(* IEC 61131-3 sources: plcassist-cli/packages/volt-lsp-iec/test-corpus/pro2193/Device/Plc Logic/Application/09 Misc/Library Manager/L_TT1P_TechnologyModules (part 2) *)

(* ---- _TM_STACKERCRANEAXISCONTROLBASE.fb ---- *)
FUNCTION_BLOCK _TM_STACKERCRANEAXISCONTROLBASE EXTENDS _TM_MotionControl
VAR_OUTPUT
	PPAR : POINTER TO _scPar_TM_StackerCraneAxisControlBase;
	PSF : POINTER TO _scSF_TM_StackerCraneAxisControlBase;
	PAP : POINTER TO _scAP_TM_StackerCraneAxisControlBase;
END_VAR
VAR_IN_OUT
	AXIS : AXIS_REF;
	DATABUSIN : ITF_DataBus;
	EADDRESS : L_TT1P_StackerCraneAddress;
	LROVERRIDE : LREAL;
	XEXECUTEBRAKETEST : BOOL;
	XEXECUTEBRAKEGRINDIN : BOOL;
	XOSCCOMP : BOOL;
	LROSCCOMPPOSSCALED : LREAL;
	LROSCCOMPLOADSCALED : LREAL;
	LRACTPOS : LREAL;
	LRACTVEL : LREAL;
	XOSCCOMPACTIVE : BOOL;
	XINPOSITION : BOOL;
	XAXISREADY : BOOL;
	ECONTROLMODE : L_MC1P_ControlMode;
	XCOMMANDABORTED : BOOL;
END_VAR
VAR
	XREGULATORONINTERNAL : BOOL;
	ETMSTATE_EXITSELECTMODE : L_TT1P_States;
	XOSCCOMP_INT : BOOL;
	XOSCCOMP_OLD : BOOL;
	XEXECUTEBRAKETEST_INT : BOOL;
	XEXECUTEBRAKEGRINDIN_INT : BOOL;
	LROVERRIDE_INT : LREAL := 1;
	LRMASTERTASKCYCLETIME : LREAL;
	LRTASKCYCLETIME : LREAL;
	SCPAR_INT : _scPar_TM_StackerCraneAxisControlBase;
	EADDRESS_INT : L_TT1P_StackerCraneAddress;
	XCOMMANDABORTED_INT : BOOL;
	XDONEBRAKEGRINDIN : BOOL;
	XDONEBRAKETEST : BOOL;
	XBRAKEFUNKTIONBUSY : BOOL;
	XSTOPACTIVE_INT : BOOL;
	XJOGGINGACTIVE_INT : BOOL;
	XHOMINGACTIVE_INT : BOOL;
	XPROFILEXYBUSY_INT : BOOL;
	XPOSITIONINGBUSY_INT : BOOL;
	XPOSITIONINGDONE_INT : BOOL;
	XBRAKETESTACTIVE : BOOL;
	XBRAKEGRINDINACTIVE : BOOL;
	XOSCCOMPENABLE_INT : BOOL;
	XOSCCOMPENABLE_OLD : BOOL;
	LRTIMECOUTERCONSTANTTORQUEVALID : LREAL;
	XSTARTCONSTANTTORQUEVALID_INT : BOOL;
	LRSTARTCONSTANTTORQUE_INT : LREAL;
	LROSCCOMPPOSSCALED_INT : LREAL := 0;
	LROSCCOMPLOADSCALED_INT : LREAL := 0;
	XOSCCOMPENABLE_LOCK : BOOL;
	LROSCCOMPPOSSCALED_LOCK : LREAL;
	LROSCCOMPLOADSCALED_LOCK : LREAL;
	XUPDATEOSCCOMPPARAMETER : BOOL;
	XAMPRATIOVALID : BOOL;
	XEIGENFREQVALID : BOOL;
	WREQUESTSOSCCOMPPARMAVALID : WORD;
	WREQUESTSOSCCOMPPARMAVALID_OLD : WORD;
	XREQUESTSOSCCOMPPARMA : BOOL;
	WRTRIGOSCCOMPPARMAVALID : WORD;
	WFTRIGOSCCOMPPARMAVALID : WORD;
	XSWLIMITDISABLED : BOOL;
	XSELECTCSVACTIVE_INT : BOOL;
	XSELECTCSPACTIVE_INT : BOOL;
	XSELECTCSPBLOKEDBYOSCCOMP : BOOL;
	EAXISSTATE_OLD : L_MC1P_AXIS_STATE;
	XPOSITIONINGDONE_OLD : BOOL;
	XAXISENABLED_OLD : BOOL;
	IFOR : INT;
	XWAITNEXTCYCLEFORSETCONTROLERMODE : BOOL;
	XINPOSITIONVALID : BOOL;
	XINPOSITION_INT : BOOL;
	LRTARGETACTPOSITION : LREAL;
	LRTARGETSETPOSITION : LREAL;
	LRPOSINWINDOW : LREAL;
	LRTIMEPOSINWINDOW : LREAL := 50;
	LRACTTIMEPOSINWINDOW : LREAL;
	XHOLDPOWEROFF_INT : BOOL;
	XDISABLEAXIS_INT : BOOL;
	XDISABLEAXIS_OLD : BOOL;
	XAXISDISABLED_INT : BOOL;
	XAXISDISABLED_OLD : BOOL;
	LRTIMECOUNTER_INT : LREAL;
	WCOUNTERAXISENABLED_INT : WORD;
	WBRAKETESTMODE : WORD;
	WBRAKETESTSTEPPER : WORD;
	WBRAKEGRINDINSTEPPER : WORD;
	LRBRAKETESTCONSTANTTORQUE : LREAL;
	LRTIMECOUNTER : LREAL;
	LRTIMEBRAKERELEASE : LREAL := 0.2;
	LRTIMEIDENTTORQUE : LREAL := 0.8;
	XRESETFILTERSTANDSTILLTORQUE : BOOL;
	WBRAKEGRINDINCYCLES_INT : WORD;
	EADDRESS_LOCK : L_TT1P_StackerCraneAddress;
	XADDRESS_LOCK : BOOL;
	ECONTROLMODECAMEFROM : L_MC1P_ControlMode;
	PELEMENT : POINTER TO L_MB1P_ChannelElement;
	PRIGHT : POINTER TO L_MB1P_ChannelElement;
	PLEFT : POINTER TO L_MB1P_ChannelElement;
	PDATA : POINTER TO L_MB1P_ChannelData;
	PDATACONTROL : POINTER TO L_MB1P_ChannelData;
	PLIST : POINTER TO L_MB1P_ListControl;
	COMIN_XLOCKCOMCHANNEL : BOOL;
	COM_XENABLE : BOOL;
	COMIN_XRESETERROR_INT : BOOL;
	COMIN_XREGULATORON_INT : BOOL;
	COMIN_XSTOP_INT : BOOL;
	COMOUTTMP_WERRORID : WORD;
	COMOUTTMP_DWERRORID : DWORD;
	COMOUT_WERRORIDSTEPPER : DWORD;
	COMOUT_DWPARSTEPPER : DWORD;
	COMOUT_DWVARSTEPPER : DWORD;
	COMOUT_DWDRIVEERRORID : DWORD;
	COMOUT_XEXECUTEMOVEXY : BOOL;
	COMOUT_XEXECUTEMOVEXY_OLD : BOOL;
	WMOVEXYEXECUTESTATE : WORD;
	COMIN_XEXECUTEPROFILEXY : BOOL;
	COMIN_XMOVEXYACTIVE : BOOL;
	COMIN_XMOVEXYBUSY : BOOL;
	COMIN_XMOVEXYDONE : BOOL;
	COMIN_XMOVEXYACTIVE_OLD : BOOL;
	COMIN_XMOVEXYDONE_OLD : BOOL;
	COMIN_XMAINTENANCEMODE : BOOL;
	COMIN_XMOVEXYCOMMANDABORT : BOOL;
	COMIN_EMASTERSTATE : WORD;
	COMIN_LRSETPOSDIST : LREAL;
	COMIN_XRESETHOLDPOWEROFF : BOOL;
	FB_COMCHANNEL : L_MB1P_ComChannelSlaveState;
	XCOMMUNICATIONVALID_LOCK : BOOL;
	XERRORCOMMUNICATION : BOOL;
	XCOMMUNICATIONVALID : BOOL;
	_XCOMERRORINVALIDMASTERCONTROLMODUL : BOOL;
	_XCOMERROR : BOOL;
	_ECOMERRORID : L_IE1P_Error;
	XERROR_INVALIDSWLIMIT : BOOL;
	XERROR_INVALIDINVERTER : BOOL;
	XERROR_NOVALIDACCELERATION_MOVEABSOLUTE : BOOL;
	XERROR_INVALIDINPUT_BRAKEGRINDIN : BOOL;
	XERROR_AXISDISABLEDISREQUIRED : BOOL;
	XWARNINGCOMMUNICATION : BOOL;
	XWARNING_INVALIDINVERTER : BOOL;
	XWARNING_AXISDISABLEDISREQUIRED : BOOL;
	FB_FILTERACTSTANDSTILLTORQUE : L_USPP_PT1Filter;
	FB_FILTERACTTORQUE : L_USPP_PT1Filter;
	FB_OSCILLATIONCOMP : L_CT1P_OscillationComp;
	FB_CALCOSCILATIONCOMPPARAMETER : L_MB1P_CalcOscilationCompParameter;
	FB_SETCONTROLLERMODE : L_MC1P_SetControlMode;
	FB_BRAKETEST : L_MC1P_BrakeTest;
	FB_BRAKEGRINDIN : L_MC1P_BrakeGrindIn;
	FB_READMACHINEDATA : L_MC1P_ReadMachineData;
	FB_DISABLESWLIMIT : L_MC1P_DisableSWLimit;
	FB_WRITEBOOLPARAMETER : MC_WriteBoolParameter;
	MC_READPARAMETERPOSINWINDOW : MC_ReadParameter := STRUCT(ParameterNumber := 130);
	MC_READPARAMETERTIMEPOSINWINDOW : MC_ReadParameter := STRUCT(ParameterNumber := 131);
	FB_RESETFOLLOWINGERROR : L_MC1P_ResetFollowingError;
	MC_READPARAMETEREXTPOSITINCNTRL : MC_ReadParameter := STRUCT(ParameterNumber := 90);
	IPARFRAME : INT;
	IMAINFRAME : INT;
	IVISUTABLESETPOS : INT := 1;
END_VAR
END_FUNCTION_BLOCK

METHOD CALL_ABC
END_METHOD

METHOD CALL_ABCCTRLREQACTIVE : BOOL
END_METHOD

METHOD CALL_ABCGENERALSETTINGS
END_METHOD

METHOD CALL_ALLOCPOINTADR
END_METHOD

METHOD CALL_COMIN
END_METHOD

METHOD CALL_COMOUT
END_METHOD

METHOD CALL_CTRLREQACTIVE : BOOL
END_METHOD

METHOD CALL_ERRORHANDLER
END_METHOD

METHOD CALL_FBMETHODS
END_METHOD

METHOD CALL_FB_BRAKEGRINDIN
END_METHOD

METHOD CALL_FB_BRAKEGRINDIN_INPUT
END_METHOD

METHOD CALL_FB_BRAKETEST
END_METHOD

METHOD CALL_FB_BRAKETEST_INPUT
END_METHOD

METHOD CALL_FB_CALCOSCILATIONCOMPPARAMETER
END_METHOD

METHOD CALL_FB_CALCOSCILATIONCOMPPARAMETER_INPUT
END_METHOD

METHOD CALL_FB_COMCHANNEL
END_METHOD

METHOD CALL_FB_DISABLESWLIMIT
END_METHOD

METHOD CALL_FB_FILTERACTTORQUE
END_METHOD

METHOD CALL_FB_OSCILLATIONCOMP
END_METHOD

METHOD CALL_FB_OSCILLATIONCOMP_INPUT
END_METHOD

METHOD CALL_FB_READPARAMETERINPOSITION
END_METHOD

METHOD CALL_FB_RESETFOLLOWINGERROR
END_METHOD

METHOD CALL_FB_SETCONTROLLERMODE
END_METHOD

METHOD CALL_FB_WRITEBOOLPARAMETER
END_METHOD

METHOD CALL_INPOSITION
END_METHOD

METHOD CALL_INITDONE
END_METHOD

METHOD CALL_INITROUTINE
END_METHOD

METHOD CALL_INTERNALCTRL
END_METHOD

METHOD CALL_MOVEXYEXECUTE
END_METHOD

METHOD CALL_OUTPUT
END_METHOD

METHOD CALL_OUTPUT_SF
END_METHOD

METHOD CALL_REQUESTS_EXT
END_METHOD

METHOD CALL_RESETCOMMANDS
END_METHOD

METHOD CALL_RESETOUTPUT
END_METHOD

METHOD CALL_RESETWARNINGS
END_METHOD

METHOD CALL_STATEMACHINE
END_METHOD

METHOD CALL_STOP
END_METHOD

METHOD GET_ADDRESS : WORD
VAR_INPUT
	IELEMENTID : INT;
	EADDRESS : L_TT1P_StackerCraneAddress;
END_VAR
END_METHOD

METHOD CALL_S000_CYCLIC
END_METHOD

METHOD CALL_S002_READY
END_METHOD

METHOD CALL_S003_HOMING
END_METHOD

METHOD CALL_S010_JOGGING
END_METHOD

METHOD CALL_S014_MOVE_ABS
END_METHOD

METHOD CALL_S060_SELECTMODECSV
END_METHOD

METHOD CALL_S123_SELECTMODECSP
END_METHOD

METHOD CALL_S186_MOVE_XY
END_METHOD

METHOD CALL_S187_MAINTENANCE
END_METHOD

METHOD CALL_S188_BRAKETEST
END_METHOD

METHOD CALL_S189_BRAKEGRINDIN
END_METHOD

METHOD CALL_S996_STOP
END_METHOD

METHOD CALL_S999_ERROR
END_METHOD

METHOD CALL_T000_ALLSTATES
END_METHOD

METHOD CALL_T002_READY
END_METHOD

(* ---- _TM_STACKERCRANEHEADCONTROLBASE.fb ---- *)
FUNCTION_BLOCK _TM_STACKERCRANEHEADCONTROLBASE EXTENDS _TM_MotionControlBase
VAR_OUTPUT
	PPAR : POINTER TO _scPar_TM_StackerCraneHeadControlBase;
	PSF : POINTER TO _scSF_TM_StackerCraneHeadControlBase;
	PAP : POINTER TO _scAP_TM_StackerCraneHeadControlBase;
END_VAR
VAR_IN_OUT
	XRESETERROR : BOOL;
	XSTOPALL : BOOL;
	SCPAR : _scPar_TM_StackerCraneHeadControlBase;
	XEXECUTEPROFILEX : BOOL;
	XEXECUTEPROFILEY : BOOL;
	XMAINTENANCEMODE : BOOL;
	DATABUSOUT : ITF_DataBus;
	XAXESREADY : BOOL;
	XAXESENABLED : BOOL;
	SCSIGNALFLOW : _scSF_TM_StackerCraneHeadControlBase;
	XAXESHOMED : BOOL;
	XPROFILEXDONE : BOOL;
	XPROFILEYDONE : BOOL;
	XPROFILEXBUSY : BOOL;
	XPROFILEYBUSY : BOOL;
	XERROR : BOOL;
	XWARNING : BOOL;
	EERRORID : L_IE1P_Error;
	ASCERRORINFO : ARRAY [1..6] OF L_TT1P_scErrorInfo;
END_VAR
VAR
	AXDONENEXTCYCLE_INT : ARRAY [1..2] OF BOOL;
	ADWREQUESTSINFOCOMIN : ARRAY [1..2] OF DWORD;
	ADWREQUESTSINFOCOMIN_OLD : ARRAY [1..2] OF DWORD;
	ADWFTRIGCOMIN : ARRAY [1..2] OF DWORD;
	ADWRTRIGCOMIN : ARRAY [1..2] OF DWORD;
	LRMASTERTASKCYCLETIME : LREAL;
	LRTASKCYCLETIME : LREAL;
	SCPAR_INT : _scPar_TM_StackerCraneHeadControlBase;
	XEXECUTEPROFILEX_INT : BOOL;
	XEXECUTEPROFILEY_INT : BOOL;
	XSTOPALL_INT : BOOL;
	XMAINTENANCEMODE_INT : BOOL;
	AXPOSITIONINGDONE_INT : ARRAY [1..2] OF BOOL;
	XPOSITIONINGDONE_INT : BOOL;
	XPOSITIONINGBUSY_INT : BOOL;
	IWAITTASKCYCLESFROSTATUSFORMCOM_INT : LREAL := 100;
	AICOUNTTASKCYCLES_INT : ARRAY [1..c_iNumOfAxisModule] OF INT;
	XXYCONTROLLERWAITSTARTX_INT : BOOL;
	XXYCONTROLLERWAITSTARTY_INT : BOOL;
	XCOMMUNICATIONVALID : BOOL;
	XLOCKCOMCHANNEL : BOOL;
	IFOR : INT;
	IDX1 : INT;
	WTEMP : WORD;
	DWTEMP : DWORD;
	DWTEMP1 : DWORD;
	DWSTATUSWORDTEMP : DWORD;
	COMIN_AXISIDX : INT;
	XWAITSTARTX_OLD : BOOL;
	XWAITSTARTY_OLD : BOOL;
	XPROFILEEXECUTE1X_OLD : BOOL;
	XPROFILEEXECUTE1Y_OLD : BOOL;
	XPROFILEEXECUTE2X_OLD : BOOL;
	XPROFILEEXECUTE2Y_OLD : BOOL;
	PLIST : POINTER TO L_MB1P_ListControl;
	PELEMENT : POINTER TO L_MB1P_ChannelElement;
	PDATA : POINTER TO L_MB1P_ChannelData;
	PDATA_AXISX : POINTER TO L_MB1P_ChannelData;
	PDATA_AXISY : POINTER TO L_MB1P_ChannelData;
	PRIGHT : POINTER TO L_MB1P_ChannelElement;
	PLEFT : POINTER TO L_MB1P_ChannelElement;
	COM_XENABLE : BOOL;
	COMIN_INUMOFAXES : INT;
	COMIN_XLOCKCOMCHANNEL : BOOL;
	COMIN_XXAXISCONTROLAVAILABLE : BOOL;
	COMIN_XYAXISCONTROLAVAILABLE : BOOL;
	COMIN_XAPAXISCONTROLAVAILABLE : BOOL;
	COMIN_XSLAVEXAXISCONTROLAVAILABLE : BOOL;
	COMIN_XSLAVEYAXISCONTROLAVAILABLE : BOOL;
	COMIN_XPOINTERTOXAXISVALID : BOOL;
	COMIN_AWPARVALIDMASK : ARRAY [1..6] OF WORD;
	COMIN_AXAXISVALID : ARRAY [1..c_iNumOfAxisModule] OF BOOL;
	COMIN_XAXESENABLED : BOOL;
	COMIN_XAXESREADY : BOOL;
	COMIN_XAXESHOMED : BOOL;
	COMIN_XSTOP : BOOL;
	COMIN_AXAXISREADY : ARRAY [1..c_iNumOfAxisModule] OF BOOL;
	COMIN_AXAXISENABLED : ARRAY [1..c_iNumOfAxisModule] OF BOOL;
	COMIN_AXHOMINGBUSY : ARRAY [1..c_iNumOfAxisModule] OF BOOL;
	COMIN_AXISHOMED : ARRAY [1..c_iNumOfAxisModule] OF BOOL;
	COMIN_AXSTOPACTIVE : ARRAY [1..c_iNumOfAxisModule] OF BOOL;
	COMIN_AXERROR : ARRAY [1..c_iNumOfAxisModule] OF BOOL;
	COMIN_AXWARNING : ARRAY [1..c_iNumOfAxisModule] OF BOOL;
	COMIN_AXABCCTRLREQACTIVE : ARRAY [1..c_iNumOfAxisModule] OF BOOL;
	COMIN_AXINPOSITION : ARRAY [1..c_iNumOfAxisModule] OF BOOL;
	COMIN_AETMSTATE : ARRAY [1..c_iNumOfAxisModule] OF WORD;
	COMIN_EERRORID : WORD;
	COMIN_AEERRORID : ARRAY [1..c_iNumOfAxisModule] OF WORD;
	COMIN_ASCERRORINFO : ARRAY [1..c_iNumOfAxisModule] OF L_TT1P_scErrorInfo;
	COMIN_AXXYPROFILEBUSY : ARRAY [1..c_iNumOfAxisModule] OF BOOL;
	COMIN_AXPOSITIONINGBUSY : ARRAY [1..c_iNumOfAxisModule] OF BOOL;
	COMIN_AXPOSITIONINGDONE : ARRAY [1..c_iNumOfAxisModule] OF BOOL;
	COMIN_ASCMINLIMITS : ARRAY [1..c_iNumOfAxisModule] OF L_TT1P_XYLimits;
	COMIN_ALRBUFFERPOSITIONNEG : ARRAY [1..c_iNumOfAxisModule] OF LREAL;
	COMIN_ALRBUFFERPOSITIONPOS : ARRAY [1..c_iNumOfAxisModule] OF LREAL;
	COMIN_ALRBUFFERVELNEG : ARRAY [1..c_iNumOfAxisModule] OF LREAL;
	COMIN_ALRBUFFERVELPOS : ARRAY [1..c_iNumOfAxisModule] OF LREAL;
	COMIN_AXBUFFERRANGE : ARRAY [1..c_iNumOfAxisModule] OF BOOL;
	COMIN_AXEXECUTEMOVEXY : ARRAY [1..c_iNumOfAxisModule] OF BOOL;
	COMIN_AXEXECUTEMOVEXY_OLD : ARRAY [1..c_iNumOfAxisModule] OF BOOL;
	COMIN_AXHOLDPOWEROFF : ARRAY [1..c_iNumOfAxisModule] OF BOOL;
	COMIN_AXPAXISVALID : ARRAY [1..c_iNumOfAxisModule] OF BOOL;
	COMIN_APAXIS : ARRAY [1..c_iNumOfAxisModule] OF POINTER TO AXIS_REF;
	COMOUT_AXRESETHOLDPOWEROFF : ARRAY [1..c_iNumOfAxisModule] OF BOOL;
	COMIN_AXOSCACTIVE : ARRAY [1..c_iNumOfAxisModule] OF BOOL;
	COMIN_AXBRAKETESTBUSY : ARRAY [1..c_iNumOfAxisModule] OF BOOL;
	COMIN_AXBRAKETESTDONE : ARRAY [1..c_iNumOfAxisModule] OF BOOL;
	COMIN_AXBRAKEGRINDINBUSY : ARRAY [1..c_iNumOfAxisModule] OF BOOL;
	COMIN_AXBRAKEGRINDINDONE : ARRAY [1..c_iNumOfAxisModule] OF BOOL;
	COMOUT_XEXECUTEPROFILEX_INT : BOOL;
	COMOUT_XEXECUTEPROFILEY_INT : BOOL;
	FB_COMCHANNEL : L_MB1P_ComChannelState;
	COMIN_XERROR_NOSTACKERCRANEAXIS : BOOL;
	XCOMMUNICATIONVALID_LOCK : BOOL;
	XERRORCOMMUNICATION : BOOL;
	_XCOMERRORINVALIDMASTERCONTROLMODUL : BOOL;
	_XCOMERROR : BOOL;
	_ECOMERRORID : L_IE1P_Error;
	XERRORDUPLICATEDADDRESS : BOOL;
	XWARNINGCOMMUNICATION : BOOL;
	XWARNING_EXECUTEXNOTPOSSIBLE : BOOL;
	XWARNING_EXECUTEYNOTPOSSIBLE : BOOL;
	XWARNING_XAXISINSERVICE : BOOL;
	XWARNING_YAXISINSERVICE : BOOL;
	XWARNING_XAXISENABLEDREQUIRED : BOOL;
	XWARNING_YAXISENABLEDREQUIRED : BOOL;
	PXAXIS : POINTER TO AXIS_REF;
	PYAXIS : POINTER TO AXIS_REF;
	XEXECUTEX_INT : BOOL;
	XEXECUTEY_INT : BOOL;
	XXYCONTROLLER_REEXECUTEX : BOOL;
	XXYCONTROLLER_REEXECUTEY : BOOL;
	EPROFILEMODEX_INT : L_TT1P_XYProfileMode;
	EPROFILEMODEY_INT : L_TT1P_XYProfileMode;
	FB_XYCONTROLLER : L_TF1P_XYController;
	IPARFRAME : INT;
	IMAINFRAME : INT;
	IVISUSELECTAXIS : INT := 1;
	ASTVISUSELECTAXIS : ARRAY [0..6] OF STRING := ['no axis selected', 'AxisX', 'AxisY', 'SlaveAxisX', 'SlaveAxisY', 'AntiPendlum', 'free axis'];
	C_INUMOFAXISMODULE : INT := 6;
END_VAR
END_FUNCTION_BLOCK

METHOD CALL_ABCCTRLREQACTIVE : BOOL
END_METHOD

METHOD CALL_ALLOCPOINTADR
END_METHOD

METHOD CALL_CHECKREQUESTS
END_METHOD

METHOD CALL_COMCHANNEL_MOVEXY
END_METHOD

METHOD CALL_COMIN
END_METHOD

METHOD CALL_COMOUT
END_METHOD

METHOD CALL_COMOUT_XYCONTROLLER_EXECUTE
END_METHOD

METHOD CALL_ERRORHANDLER
END_METHOD

METHOD CALL_ERRORHANDLER_SCERRORINFO
END_METHOD

METHOD CALL_FBMETHODS
END_METHOD

METHOD CALL_FB_COMCHANNEL
END_METHOD

METHOD CALL_FB_XYCONTROLLER
END_METHOD

METHOD CALL_FB_XYCONTROLLER_INPUT
END_METHOD

METHOD CALL_INITDONE
END_METHOD

METHOD CALL_INITROUTINE
END_METHOD

METHOD CALL_INTERNALCTRL
END_METHOD

METHOD CALL_OUTPUT
END_METHOD

METHOD CALL_OUTPUT_SF
END_METHOD

METHOD CALL_REQUESTS_COMIN
END_METHOD

METHOD CALL_REQUESTS_EXT
END_METHOD

METHOD CALL_RESETCOMMANDS
END_METHOD

METHOD CALL_RESETCOUNTER
END_METHOD

METHOD CALL_RESETOUTPUT
END_METHOD

METHOD CALL_RESETWARNINGS
END_METHOD

METHOD CALL_STATEMACHINE
END_METHOD

METHOD CALL_TMFUNCTIONALITY
END_METHOD

METHOD CALL_S000_CYCLIC
END_METHOD

METHOD CALL_S002_READY
END_METHOD

METHOD CALL_S186_MOVE_XY
END_METHOD

METHOD CALL_S187_MAINTENANCE
END_METHOD

METHOD CALL_S996_STOP
END_METHOD

METHOD CALL_S998_SERVICE
END_METHOD

METHOD CALL_S999_ERROR
END_METHOD

METHOD CALL_T000_ALLSTATES
END_METHOD

METHOD CALL_T002_READY
END_METHOD

(* ---- _TM_TABLEPOSITIONINGBASE.fb ---- *)
FUNCTION_BLOCK _TM_TABLEPOSITIONINGBASE EXTENDS _TM_MotionControl
VAR_OUTPUT
	PPAR : POINTER TO _scPar_TM_TablePositioningHigh;
	PSF : POINTER TO _scSF_TM_TablePositioningHigh;
	PAP : POINTER TO _scSF_TM_TablePositioningHigh;
END_VAR
VAR_IN_OUT
	AXIS : AXIS_REF;
	XRESETHOMEPOSITION : BOOL;
	XHWLIMITPOS : BOOL;
	XHWLIMITNEG : BOOL;
	XEXECUTEPOSITIONING : BOOL;
	XABORTPOSITIONING : BOOL;
	XFINISHPOSITIONING : BOOL;
	EPROFILENUMBER : L_TT1P_ProfileNumber;
	XTPRECEIVE : BOOL;
	LRACTTPPOSITION : LREAL;
	LRCYCPOSEXTENCODER : LREAL;
	LRSETTORQUELIMITPOS : LREAL;
	LRSETTORQUELIMITNEG : LREAL;
	LRSETOVERRIDEVELOCITY : LREAL;
	LRSETOVERRIDEACCDEC : LREAL;
	LRSETOVERRIDEJERK : LREAL;
	XPOSITIONINGACTIVE : BOOL;
	XPOSITIONINGDONE : BOOL;
	XDRIVEINTARGET : BOOL;
	LRACTPOS : LREAL;
	LRACTVEL : LREAL;
	LRACTFOLLOWINGERROR : LREAL;
	XTPRECEIVED : BOOL;
	XTPMISSED : BOOL;
	XTPOUTOFWINDOW : BOOL;
	EACTIVEPROFILE : L_TT1P_ProfileNumber;
END_VAR
VAR
	SCPAR_INT : _scPar_TM_TablePositioningHigh;
	XEXECUTEPOSITIONING_INT : BOOL;
	XABORTPOSITIONING_INT : BOOL;
	XFINISHPOSITIONING_INT : BOOL;
	XAUTOMATICUPDATE_INT : BOOL;
	LRACTTPPOSITION_INT : LREAL;
	EPROFILENUMBER_INT : L_TT1P_ProfileNumber;
	LRSETTORQUELIMITPOS_INT : LREAL;
	LRSETTORQUELIMITNEG_INT : LREAL;
	LRSETOVERRIDEVELOCITY_INT : LREAL;
	LRSETOVERRIDEACCDEC_INT : LREAL;
	LRSETOVERRIDEJERK_INT : LREAL;
	XRESETHOMEPOSITION_INT : BOOL;
	XHWLIMITPOS_INT : BOOL;
	XHWLIMITNEG_INT : BOOL;
	XTPRECEIVED_INT : BOOL;
	XTPMISSED_INT : BOOL;
	XTPOUTOFWINDOW_INT : BOOL := FALSE;
	XPOSITIONINGACTIVE_INT : BOOL;
	XPOSITIONINGDONE_INT : BOOL;
	XTPRECEIVE_INT : BOOL := FALSE;
	BYSTEPPER : BYTE;
	WSEQUENCEPROFILE : WORD := 0;
	XSEQUENCEPROFILEACTIVE : BOOL;
	XPOSDISABLEFOLLOWPROFILE : BOOL;
	LRSETPOSSEQUENCEPROFILE : LREAL;
	LRSETPOSFINISHTARGET : LREAL;
	LRFINALPOSITION : LREAL;
	XINTARGET : BOOL;
	XHOMINGEXECUTEOLD_INT : BOOL;
	HWLIMITSWITCHINTERFACE : L_MC1P_HWLimitSwitchInterface;
	RESETHOMEPOSITION : L_MC1P_ResetHomePosition;
	SMC_MOVECONTINUOUSABSOLUTE : MC_MoveContinuousAbsolute;
	SMC_MOVECONTINUOUSRELATIVE : MC_MoveContinuousRelative;
	TORQUELIMITS : L_MC1P_SetTorqueLimit;
	MC_HALT : MC_Halt;
	CONVERTTP : L_MB1P_TpConvertTp;
	READWINDOWPARAMETER : MC_ReadParameter;
	LRTARGETDISTANCE_INT : LREAL := 0;
	XPOSITIONINGABORTED_INT : BOOL := FALSE;
	XTPINSIDEWINDOW : BOOL := FALSE;
	LRTPPOSITIONINGTARGET : LREAL;
	LRACTUALPROFILEDISTANCE : LREAL;
	LRPOSITIONOLD : LREAL;
	XRESTARTPROFILE : BOOL;
	WCOUNTER : WORD;
	XEXECUTEOLD : BOOL;
	LRVELOCITYOLD : LREAL;
	XSTARTPROFILEOLD : BOOL;
	XRESTARTVELPROFILE : BOOL;
	XERRORTRAVERSIONRANGE : BOOL := FALSE;
	XNOPROFILESELECTED : BOOL := FALSE;
	XPOSITIONINGMODEINVALID : BOOL := FALSE;
	XAXISNOTHOMED : BOOL := FALSE;
	XTPRECEIVEOLD : BOOL := FALSE;
	EABORTEDPROFILE : L_TT1P_ProfileNumber;
	XTPWINDOWOPEN : BOOL;
	LRFINALPOSITIONMODULO : LREAL;
	XVISPOINTMIN : BOOL;
	XVISPOINTMAX : BOOL;
	XVISUSETPOSUP : BOOL;
	XVISUSETPOSDOWN : BOOL;
	RTRIGUP : R_TRIG;
	RTRIGDOWN : R_TRIG;
	IMAXPOINTS : INT := 13;
	IPOINT : INT := 1;
	LRTARGETWINDOW : LREAL;
	XINSIDEWINDOWFLAG : BOOL;
	XTPOUTSIDEWINDOW_TPMETHOD : BOOL;
	XTPINSIDEWINDOW_TPMETHOD : BOOL;
	LRACTUALSEQUENCESTARTPOSITION : LREAL;
	XPROFILECHAININGWITHVELOCITY : BOOL;
	XTPOUTSIDEOFWINDOW : BOOL := FALSE;
	PXMOVEFUNBUSY : POINTER TO BOOL;
	ISTATESTEPPER : INT := 0;
	XFIRSTPOSITIONINGCYCLE : BOOL := TRUE;
	XAXISVIRTUAL : BOOL := FALSE;
	XINENDVELOCITY : BOOL := FALSE;
	XTPPROFILEACTIVE : BOOL;
	XTPDURINGPOSITIONING : BOOL := FALSE;
	XPOSITIVEPROFILEVELOCITY : BOOL;
	XABORTACTIVE_INT : BOOL;
	XFINISHINGPOSITIONING_INT : BOOL;
	XEXECUTEPOSITIONINGFLAG : BOOL;
	XFINISHPOSITIONINGFLAG : BOOL;
	XABSOLUTEINENDVELOCITYOLD : BOOL;
	XRELATIVEINENDVELOCITYOLD : BOOL;
	XFUNDONEOLD : BOOL;
	XINPOSITIONOLD : BOOL;
	XFUNBUSYOLD : BOOL := FALSE;
	XPOSITIONINGDONEACTIVE : BOOL := FALSE;
	XABORTBUSYOLD : BOOL := FALSE;
	LRSETPOSITIONOLD : LREAL;
	XLASTPROFILE : BOOL;
	XCINHNOERROR : BOOL := FALSE;
	LRMODULOTARGETPOS : LREAL := 0;
	LRDIFFINSIDECYCLE : LREAL := 0;
	LRINTEGRATOR : LREAL;
	XINTEGRATORACTIVE : BOOL;
	XMOVERELEXECUTEOLD : BOOL;
	XEXECUTEMOVECONTINUOUSOLD : BOOL;
	XFIRSTSTARTRELATIVEPROFILE : BOOL;
END_VAR
END_FUNCTION_BLOCK

METHOD CALL_MC_SETTORQUE_INPUT
END_METHOD

METHOD CALL_ALLOCPOINTADR
END_METHOD

METHOD CALL_ERRORHANDLER
END_METHOD

METHOD CALL_FBMETHODS
END_METHOD

METHOD CALL_FBS
END_METHOD

METHOD CALL_FIRSTCYCLE
END_METHOD

METHOD CALL_INITDONE
END_METHOD

METHOD CALL_INITROUTINE
END_METHOD

METHOD CALL_INTERNALCTRL
END_METHOD

METHOD CALL_MC1P_HWLIMITSWITCH
END_METHOD

METHOD CALL_MC1P_RESETHOMEPOSITION
END_METHOD

METHOD CALL_OUTPUT
END_METHOD

METHOD CALL_READPOSITIONINGWINDOW
END_METHOD

METHOD CALL_REQUESTS_EXT
END_METHOD

METHOD CALL_RESETCOMMANDS
END_METHOD

METHOD CALL_RESETOUTPUTS
END_METHOD

METHOD CALL_STATEMACHINE
END_METHOD

METHOD CALL_TOUCHPROBESOURCE
END_METHOD

METHOD CALL_TPWINDOWSTATUS
END_METHOD

METHOD CALL_VISUPROFILES
END_METHOD

METHOD CALL_ABC
END_METHOD

METHOD CALL_020_RELATIVEENTRY
END_METHOD

METHOD CALL_022_RELATIVEFINALVELOCITY
END_METHOD

METHOD CALL_024_RELATIVE
END_METHOD

METHOD CALL_02_STARTSEQUENCEPROFILES
END_METHOD

METHOD CALL_110_ABORTPOSITIONING
END_METHOD

METHOD CALL_200_ERROR
END_METHOD

METHOD CALL_90_SEQUENCEPROFILE
END_METHOD

METHOD CALL_S000_CYCLIC
END_METHOD

METHOD CALL_S080_POSITIONING
END_METHOD

METHOD CALL_S081_POSITIONING_EXIT
END_METHOD

METHOD CALL_S996_STOP
END_METHOD

METHOD CALL_S999_ERROR
END_METHOD

METHOD CALL_T002_READY
END_METHOD

(* ---- _TM_VIRTUALMASTERBASE.fb ---- *)
FUNCTION_BLOCK _TM_VIRTUALMASTERBASE EXTENDS _TM_MotionControl
VAR_OUTPUT
	PPAR : POINTER TO _scPar_TM_VirtualMasterHigh;
END_VAR
VAR_IN_OUT
	VIRTUALAXIS : AXIS_REF;
	XCONTINUOUS : BOOL;
	XCYCLE : BOOL;
	XLOADSTARTPOS : BOOL;
	LRSETVEL : LREAL;
	LRSTARTPOS : LREAL;
	LRTARGETPOS : LREAL;
	XINTARGET : BOOL;
	LRACTPOS : LREAL;
	LRACTVEL : LREAL;
	LRSETPOSOUT : LREAL;
	LRSETVELOUT : LREAL;
END_VAR
VAR
	SCPAR_INT : _scPar_TM_VirtualMasterHigh;
	XCONTINUOUS_INT : BOOL;
	XCYCLE_INT : BOOL;
	XLOADSTARTPOS_INT : BOOL;
	LRSTARTPOS_INT : LREAL;
	LRTARGETPOS_INT : LREAL;
	LRSETVEL_INT : LREAL;
	LRSETVEL_LOCK : LREAL;
	EDIRECTION_LOCK : MC_DIRECTION;
	XSYNCMASTERAXIS_INT : BOOL;
	LRMASTERSTARTDISTANCE_INT : LREAL;
	LRMASTERSYNCPOSITION_INT : LREAL;
	LRSLAVESYNCPOSITION_INT : LREAL;
	WOLDSTATE : WORD;
	XSYNCMASTERAXIS_OLD : BOOL;
	XCONTINUOUS_OLD : BOOL;
	XCYCLE_OLD : BOOL;
	XSTOP_OLD : BOOL;
	XLOADSTARTPOS_OLD : BOOL;
	XOLDENABLE : BOOL;
	XSTARTPOSOUTRANGE : BOOL;
	LRTARGETPOS_SAVE : LREAL;
	XSP_EXECUTE : BOOL;
	XSP_STARTED : BOOL;
	XMOVETOTARGETPOSACTIVE : BOOL;
	BYSTEPPERMOVETOTARGETPOS : BYTE;
	LRCYCLELENGTH : LREAL;
	XMASTERITFVALID : BOOL;
	BYMASTERID : POINTER TO BYTE;
	XMASTERITFVALID_LOCK : BOOL;
	BYMASTERID_LOCK : POINTER TO BYTE;
	EMASTERTRAVERSINGRANGE : L_MC1P_TraversingRange;
	LRMASTERCYCLELENGTH : LREAL;
	LRMASTERSETPOSITIONFORSYNC : LREAL;
	LRMASTERSETVELOCITYFORSYNC : LREAL;
	LRMASTERSETACCELERATIONFORSYNC : LREAL;
	XSYNCOUTATTARGETPOS : BOOL;
	XSYNCOUTATTARGETPOSACTIVE : BOOL;
	XINTERNALCONTR_R_EDGE : R_TRIG;
	FB_SETPOSITION : MC_SetPosition;
END_VAR
END_FUNCTION_BLOCK

METHOD CALL_ABC
END_METHOD

METHOD CALL_ALLOCPOINTADR
END_METHOD

METHOD CALL_ERRORHANDLER
END_METHOD

METHOD CALL_FBMETHODS
END_METHOD

METHOD CALL_INITROUTINE
END_METHOD

METHOD CALL_INTERNALCTRL
END_METHOD

METHOD CALL_MC_SETPOSITION
END_METHOD

METHOD CALL_MASTERAXISREF
VAR_INPUT
	MASTERAXIS : L_MC1P_IAXIS_REF_MASTERVALUES;
END_VAR
END_METHOD

METHOD CALL_OUTPUT
END_METHOD

METHOD CALL_REQUESTS_EXT
END_METHOD

METHOD CALL_RESETABCMOVEEXECUTE
END_METHOD

METHOD CALL_RESETCOMMANDS
END_METHOD

METHOD CALL_RESETOUTPUT
END_METHOD

METHOD CALL_SETABCMOVEPAR
END_METHOD

METHOD CALL_SETABCMOVESETVEL
END_METHOD

METHOD CALL_STATEMACHINE
END_METHOD

METHOD CALL_S000_CYCLIC
END_METHOD

METHOD CALL_S002_READY
END_METHOD

METHOD CALL_S035_MOVE_TO_TARGET_POS
END_METHOD

METHOD CALL_S060_CONTMOTION
END_METHOD

METHOD CALL_S130_CYCLICMOTION
END_METHOD

METHOD CALL_S999_ERROR
END_METHOD

METHOD CALL_T002_READY
END_METHOD

METHOD CALL_T035_MOVE_TO_TARGET_POS
END_METHOD

METHOD CALL_T060_CONTMOTION
END_METHOD

(* ---- _TM_VIRTUALMASTERHIGH.fb ---- *)
FUNCTION_BLOCK _TM_VIRTUALMASTERHIGH EXTENDS _TM_VirtualMasterBase
VAR_INPUT
	MASTERAXIS : L_MC1P_IAXIS_REF_MASTERVALUES;
END_VAR
VAR_IN_OUT
	XSYNCMASTERAXIS : BOOL;
	XACCDECSYNC : BOOL;
	XSYNCHRONISED : BOOL;
END_VAR
VAR
	XWARNING_SYNCMODEVELACCREQUIRED : BOOL;
	XWARNING_INVALIDSYNCSLAVEDIRECTION : BOOL;
	XERROR_INVALIDSYNCSLAVEDIRECTION : BOOL;
	BYSTEPPESYNCOUTATTARGETPOS : BYTE;
	XCONTMOTION2SYNC : BOOL;
	XMOVETARGET2CONTMOTION : BOOL;
	FB_CLUTCHEXTENDEDBASE : L_MB1P_ClutchExtendedBase;
	FB_AXISCONTROLBYPOS : L_MC1P_ControlSetValues;
END_VAR
END_FUNCTION_BLOCK

METHOD CALL_ERRORHANDLER
END_METHOD

METHOD CALL_FBMETHODS
END_METHOD

METHOD CALL_FB_AXISCONTROLBYPOS
END_METHOD

METHOD CALL_FB_CLUTCHEXTENDEDBASE
END_METHOD

METHOD CALL_INITROUTINE
END_METHOD

METHOD CALL_INTERNALCTRL
END_METHOD

METHOD CALL_INTERNALCTRLSTATE
END_METHOD

METHOD CALL_OUTPUT
END_METHOD

METHOD CALL_REQUESTS_EXT
END_METHOD

METHOD CALL_RESETCOMMANDS
END_METHOD

METHOD CALL_SETCLUTCHPOSPAR
END_METHOD

METHOD CALL_STATEMACHINE
END_METHOD

METHOD CALL_SYNCDRIVE
END_METHOD

METHOD SWITCHTOEXTMASTER
END_METHOD

METHOD CALL_S030_SYNCHRONISING_POS
END_METHOD

METHOD CALL_S031_POS_IS_SYNCHRONISED
END_METHOD

METHOD CALL_S035_MOVE_TO_TARGET_POS
END_METHOD

METHOD CALL_S060_CONTMOTION
END_METHOD

METHOD CALL_S999_ERROR
END_METHOD

METHOD CALL_T002_READY
END_METHOD

METHOD CALL_T035_MOVE_TO_TARGET_POS
END_METHOD

METHOD CALL_T060_CONTMOTION
END_METHOD

(* ---- _TM_VIRTUALMASTERSTATE.fb ---- *)
FUNCTION_BLOCK _TM_VIRTUALMASTERSTATE EXTENDS _TM_VirtualMasterBase
VAR_INPUT
	MASTERAXIS : L_MC1P_IAXIS_REF_MASTERVALUES;
END_VAR
VAR_OUTPUT
	PPARSTATE : POINTER TO _scPar_TM_VirtualMasterStateExtension;
END_VAR
VAR_IN_OUT
	XSYNCMASTERAXIS : BOOL;
	XACCDECSYNC : BOOL;
	XSYNCHRONISED : BOOL;
END_VAR
VAR
	SCPARSTATE_INT : _scPar_TM_VirtualMasterStateExtension;
	GEARIN : MC_GearIn;
END_VAR
END_FUNCTION_BLOCK

METHOD CALL_ALLOCPOINTADR
END_METHOD

METHOD CALL_ALLOCPOINTADRSTATE
END_METHOD

METHOD CALL_ERRORHANDLER
END_METHOD

METHOD CALL_FBMETHODS
END_METHOD

METHOD CALL_GEARIN
END_METHOD

METHOD CALL_INITROUTINE
END_METHOD

METHOD CALL_INTERNALCTRL
END_METHOD

METHOD CALL_INTERNALCTRLSTATE
END_METHOD

METHOD CALL_OUTPUT
END_METHOD

METHOD CALL_RESETCOMMANDS
END_METHOD

METHOD CALL_RESETOUTPUT
END_METHOD

METHOD CALL_STATEMACHINE
END_METHOD

METHOD SWITCHTOEXTMASTER
END_METHOD

METHOD CALL_S000_CYCLIC
END_METHOD

METHOD CALL_S040_SYNCHRONISING_VEL
END_METHOD

METHOD CALL_S041_VELSYNCHRONISED
END_METHOD

METHOD CALL_S999_ERROR
END_METHOD

(* ---- _TM_WINDER.fb ---- *)
FUNCTION_BLOCK _TM_WINDER EXTENDS _TM_MotionControl
VAR_IN_OUT
	AXIS : AXIS_REF;
	MATERIALCOUNTERAXIS : L_MC1P_IAXIS_REF_POOL;
	PERSISTENTVAR : L_TT1P_PersistentVarWinder;
	XMATERIALFEEDING : BOOL;
	XWINDINGDIRECTION : BOOL;
	XLOADDIAM : BOOL;
	LRSETDIAM : LREAL;
	XHOLDDIAM : BOOL;
	XDIAMCALCREDUCED : BOOL;
	XWEBBREAKMONIT : BOOL;
	XJOGLINEPOS : BOOL;
	XJOGLINENEG : BOOL;
	XTRIMLINEPOS : BOOL;
	XTRIMLINENEG : BOOL;
	XSYNCLINEVEL : BOOL;
	XTENSCURVE : BOOL;
	LRSETTENS : LREAL;
	LRSETLINEVEL : LREAL;
	XSETMATERIALCOUNTER : BOOL;
	XSYNCHRONISED : BOOL;
	XACCDECSYNC : BOOL;
	XUNWIND : BOOL;
	XWEBBREAK : BOOL;
	XHOLDDIAMACTIVE : BOOL;
	XDIAMMAX : BOOL;
	XDIAMMIN : BOOL;
	LRSETDIAMOUT : LREAL;
	LRSETDIAMSCALEDOUT : LREAL;
	LRSETLINEVELSCALEDOUT : LREAL;
	LRACTTOTALTRQSCALED : LREAL;
	LRWNDSPDREF : LREAL;
	LRMATERIALCOUNTER : LREAL;
	LRLIMITLINEVEL : LREAL;
END_VAR
VAR
	XWINDINGDIRECTION_INT : BOOL := FALSE;
	XWINDINGDIRECTIONSTANDSTILL_INT : BOOL := FALSE;
	XMATERIALFEEDING_INT : BOOL := FALSE;
	XLOADDIAM_INT : BOOL;
	LRSETDIAM_INT : LREAL;
	XHOLDDIAM_INT : BOOL;
	XDIAMCALCREDUCED_INT : BOOL;
	XWEBBREAKMONIT_INT : BOOL;
	XJOGLINEPOS_INT : BOOL;
	XJOGLINENEG_INT : BOOL;
	XTRIMLINEPOS_INT : BOOL;
	XTRIMLINENEG_INT : BOOL;
	XSYNCLINEVEL_INT : BOOL;
	LRSETTENS_INT : LREAL;
	XTENSCURVE_INT : BOOL;
	XSYNCHRONISED_INT : BOOL;
	XACCDECSYNC_INT : BOOL;
	XSETMATERIALCOUNTER_INT : BOOL;
	AP10_XSETTRQOFFSET_INT : BOOL;
	AP10_LRSETTRQOFFSET_INT : LREAL;
	AP09_XSETVELOFFSET_INT : BOOL;
	AP09_LRSETVELOFFSET_INT : LREAL;
	XLINEVELDIAMCALC_INT : BOOL;
	LRSETLINEVELDIAMCALC_INT : LREAL;
	XSYNCLINEVEL_INT_OLD : BOOL;
	XUNWIND_OLD : BOOL;
	LRSETDIAMOUT_OLD : LREAL;
	XLOADDIAM_INT_OLD : BOOL;
	XERRORINVALIDINVERTER : BOOL;
	XWARNINGAXISNOTHOMED : BOOL;
	DISETLOWERSPEEDLIMIT : DINT;
	DISETUPPERSPEEDLIMIT : DINT;
	DIOFFSETTORQUE : DINT;
	LRREFERENCEMOTORREELSPEED : LREAL := 0;
	LRREFERENCEREELSPEEDWINDER : LREAL := 0;
	LRREFERENCETORQUEWINDER : LREAL := 0;
	LRREFERENCETORQUEWINDERINV : LREAL;
	LRREFERENCEMOTORTORQUE : LREAL := 0;
	LRFEEDCONSTANT : LREAL;
	LRFEEDCONSTANT_ABS : LREAL;
	LRFEEDCONSTANTINV : LREAL;
	LRFEEDCONSTANTINV_ABS : LREAL;
	LRCYCLELENGTH_INV : LREAL;
	LRCYCLELENGTH : LREAL;
	LRGEARNUMERATOR : LREAL;
	LRGEARDENOMINATOR : LREAL;
	DWGEARNUMERATOR_LOCK : DWORD;
	DWGEARDENOMINATOR_LOCK : DWORD;
	XIDENTDIAMACTIVE_INT : BOOL;
	LRREADAXISREELSPEED : LREAL;
	LRCIRCUMFERENCE : LREAL;
	LRCIRCUMFERENCE_INV : LREAL;
	XSPEEDLIMITENABLED : BOOL;
	XDECOUPLINGLIMITREELSPEED : BOOL;
	XDCALCDISTANCEINIT : BOOL;
	WWINDERID : WORD;
	LRREELSPEEDMIN : LREAL := 0.002;
	LRMINLINEVEL : LREAL;
	LRSETWNDSPEEDUPPERLIMIT : LREAL;
	LRSETWNDSPEEDLOWERLIMIT : LREAL;
	LRSETSPEEDCTRLGAINADAPT : LREAL := 1;
	LRSETSPEEDOFFSET : LREAL := 0;
	XTRIGGERCALCDIAM : BOOL;
	XTRIGGERCALCDIAM_OLD : BOOL;
	WNUMOFAXIS : WORD;
	XMATERIALCOUNTERAXISVALID : BOOL := FALSE;
	PMATERIALCOUNTERAXIS : POINTER TO AXIS_REF;
	ETMSTATE_EXITSELECTMODE : L_TT1P_States := 2;
	ECONTROLMODECAMEFROM : L_MC1P_ControlMode;
	XWAITNEXTCYCLEFORSETCONTROLERMODE : BOOL;
	XSELECTCSVACTIVE_INT : BOOL;
	XSELECTCSPACTIVE_INT : BOOL;
	XSELECTCSTACTIVE_INT : BOOL;
	AP_XSETCONTROLLERMODE : BOOL;
	PPARWINDER : POINTER TO _scPar_TM_Winder;
	XWEBBREAKEXT : BOOL := FALSE;
	LRPICTRLINTVALUE : LREAL := 0;
	XPICTRLLOADINTVALUE : BOOL := FALSE;
	XENABLETRQFOLLOWER : BOOL;
	LRACTTOTALTORQUE : LREAL;
	LRSETTORQUEOFFSET : LREAL := 0;
	LRSETTOTALTORQUE : LREAL;
	LRSETMOTORTORQUE : LREAL;
	LRACTMOTORTORQUE : LREAL;
	LRSETTOTALVELOCITY : LREAL;
	LRVARMINERTIASCALED : LREAL;
	LRWNDVELREF : LREAL;
	LRSETPOSITION_OLD : LREAL;
	FB_READPARAMETER : MC_ReadParameter;
	FB_READMACHINEDATA : L_MC1P_ReadmachineData;
	FB_READMACHINEDATAMATCNTAXIS : L_MC1P_ReadmachineData;
	FB_FOLLOWVELOCITY : L_MC1P_FollowSetValues;
	FB_FOLLOWTORQUE : L_MC1P_SetTorqueOffset;
	FB_SETCONTROLLERMODE : L_MC1P_SetControlMode;
	FB_TORQUECONTROL : L_MC1P_TorqueControl;
	L_MB1P_CURVESETDIAMETER : L_USPP_Curve;
	L_MB1P_CALCDIAMETER1 : L_TB1P_CalcDiameter;
	L_MB1P_TENSIONCURVE1 : L_TB1P_TensionCurve;
	FB_RAMPGENERATOR1 : L_MC1P_RampGenerator;
	FB_WINDERSYNCHRONISELINE1 : L_MB1P_WinderSynchroniseLine;
	FM_WINDERJOGGING1 : L_TF1P_WinderJogging;
	WMATERIALLENGTHCOUNTERMODE : WORD;
	FB_MATERIALLENGTHCOUNTER : L_MB1P_MaterialLengthCounterFromVel;
	FB_MATERIALLENGTHCOUNTERPOS : L_MB1P_MaterialLengthCounterFromPos;
	XINVERTDIRECTION : BOOL;
	LRREELSPEEDINTEGRATE : LREAL;
	XDIAMCALCULATED_INT : BOOL;
	XINVALIDRETAIN : BOOL;
	LRSETDIAMOUTRETAIN : LREAL;
END_VAR
END_FUNCTION_BLOCK

METHOD CALL_ALLOCPOINTADR
END_METHOD

METHOD CALL_CALCCIRCUMFERENCE
END_METHOD

METHOD CALL_CTRLREQACTIVE : BOOL
END_METHOD

METHOD CALL_ERRORHANDLER
END_METHOD

METHOD CALL_FBMETHODS
END_METHOD

METHOD CALL_FBMETHODS_WND
END_METHOD

METHOD CALL_FB_MATERIALLENGTHCOUNTER
END_METHOD

METHOD CALL_FB_MATERIALLENGTHCOUNTER_INPUT
END_METHOD

METHOD CALL_FB_RAMPGENERATOR
END_METHOD

METHOD CALL_FB_RAMPGENERATOR_INPUT
END_METHOD

METHOD CALL_FB_READPARAMETER
END_METHOD

METHOD CALL_FB_READMACHINEDATA
END_METHOD

METHOD CALL_FB_READMACHINEDATAMATCNTAXIS
END_METHOD

METHOD CALL_FB_SETCONTROLLERMODE
END_METHOD

METHOD CALL_FB_TORQUECONTROL
END_METHOD

METHOD CALL_FB_WINDERSYNCHRONISELINE
END_METHOD

METHOD CALL_FB_WNDCALCDIAMETER
END_METHOD

METHOD CALL_FB_WNDCALCDIAMETER_CALCDISTACE
END_METHOD

METHOD CALL_FB_WNDCALCDIAMETER_HOLDDIAMETER
END_METHOD

METHOD CALL_FB_WNDCALCDIAMETER_INPUT
END_METHOD

METHOD CALL_FM_WINDERJOGGING
END_METHOD

METHOD CALL_FIRSTCYCLE
END_METHOD

METHOD CALL_FOLLOWTORQUE
END_METHOD

METHOD CALL_FOLLOWVELOCITY
END_METHOD

METHOD CALL_INITDONE
END_METHOD

METHOD CALL_INITROUTINE
END_METHOD

METHOD CALL_INTERNALCTRL
END_METHOD

METHOD CALL_INTERNALCTRLACTIVE
END_METHOD

METHOD CALL_INTERNALCTRLNOTACTIVE
END_METHOD

METHOD CALL_LIMITLINEVEL
END_METHOD

METHOD CALL_LIMITEDINPUT
END_METHOD

METHOD CALL_OUTPUT
END_METHOD

METHOD CALL_READACTUALTORQUE
END_METHOD

METHOD CALL_READAXISREELSPEED
END_METHOD

METHOD CALL_REQUESTS_EXT
END_METHOD

METHOD CALL_RESETCOMMANDS
END_METHOD

METHOD CALL_RESETOUTPUT
END_METHOD

METHOD CALL_RESETPERSISTENTVARWINDER
END_METHOD

METHOD CALL_RESETWARNINGS
END_METHOD

METHOD CALL_SETPERSISTENTVARWINDER
END_METHOD

METHOD CALL_SETSPEEDPOINT
END_METHOD

METHOD CALL_SETTORQUE
END_METHOD

METHOD CALL_SETWINDERID
END_METHOD

METHOD CALL_STATEMACHINE
END_METHOD

METHOD CALL_TBCURVESETDIAMETER : LREAL
END_METHOD

METHOD CALL_WNDTENSIONCURVE
END_METHOD

METHOD CALL_WNDTENSIONCURVE_INPUT
END_METHOD

METHOD CALL_ABC
END_METHOD

METHOD GET_ESTATE : L_TT1P_States
END_METHOD

METHOD GET_ETMSTATE : L_TT1P_States
END_METHOD

METHOD GET_LRACTMOTORTORQUE : LREAL
END_METHOD

METHOD GET_LRCALCDIAMDIST : LREAL
END_METHOD

METHOD GET_LRCALCDIAMLINESPEED : LREAL
END_METHOD

METHOD GET_LRCALCDIAMREELSPEED : LREAL
END_METHOD

METHOD GET_LRFEEDCONSTANT : LREAL
END_METHOD

METHOD GET_LRLOWERSPEEDLIMIT : LREAL
END_METHOD

METHOD GET_LRMOTORTORQUEREF : LREAL
END_METHOD

METHOD GET_LRREELSPEEDREF : LREAL
END_METHOD

METHOD GET_LRSETMOTORTORQUE : LREAL
END_METHOD

METHOD GET_LRSETSPEEDCTRLGAINADAPT : LREAL
END_METHOD

METHOD GET_LRSETTOTALTORQUE : LREAL
END_METHOD

METHOD GET_LRSETTOTALTRQ : LREAL
END_METHOD

METHOD GET_LRTASKCYCLE : LREAL
END_METHOD

METHOD GET_LRUPPERSPEEDLIMIT : LREAL
END_METHOD

METHOD GET_LRVARMINERTIASCALED : LREAL
END_METHOD

METHOD GET_LRWINDERTORQUEREF : LREAL
END_METHOD

METHOD GET_XCOMMUNICATION : BOOL
END_METHOD

METHOD GET_XDIAMWEBBREAKENABLE : BOOL
VAR_OUTPUT
	XUNIDIRECT : BOOL;
	XUNWINDACTIVE : BOOL;
END_VAR
END_METHOD

METHOD CALL_COUPLINGREELSPEEDLIMIT
END_METHOD

METHOD CALL_DECOUPLINGREELSPEEDLIMIT
END_METHOD

METHOD RESET_SYSTEMFAULT
END_METHOD

METHOD SET_SYSTEMFAULT
VAR_INPUT
	IN : L_IE1P_Error;
END_VAR
END_METHOD

METHOD SET_ESTATE
VAR_INPUT
	IN : L_TT1P_States;
END_VAR
END_METHOD

METHOD SET_LRFEEDCONSTANT
VAR_INPUT
	LRIN : LREAL := 0;
END_VAR
END_METHOD

METHOD SET_LRPICTRLINTVALUE
VAR_INPUT
	LRIN : LREAL := 0;
END_VAR
END_METHOD

METHOD SET_LRREFERENCEMOTORTORQUE
VAR_INPUT
	LRIN : LREAL := 0;
END_VAR
END_METHOD

METHOD SET_LRREFERENCEREELSPEED
VAR_INPUT
	LRIN : LREAL := 0;
END_VAR
END_METHOD

METHOD SET_LRSPEEDOFFSET
VAR_INPUT
	LRIN : LREAL := 0;
END_VAR
END_METHOD

METHOD SET_LRTORQUEOFFSET
VAR_INPUT
	LRIN : LREAL := 0;
END_VAR
END_METHOD

METHOD SET_XPICTRLLOADINTVALUE
VAR_INPUT
	XIN : BOOL := FALSE;
END_VAR
END_METHOD

METHOD SET_XSPEEDLIMITENABLEDEXT
VAR_INPUT
	XIN : BOOL := TRUE;
END_VAR
END_METHOD

METHOD SET_XWEBBREAK
VAR_INPUT
	XIN : BOOL := FALSE;
END_VAR
END_METHOD

METHOD CALL_S000_CYCLIC
END_METHOD

METHOD CALL_S002_READY
END_METHOD

METHOD CALL_S010_JOGGING
END_METHOD

METHOD CALL_S020_SYNCLINEVEL
END_METHOD

METHOD CALL_S060_SELECTMODECSV
END_METHOD

METHOD CALL_S070_SELECTMODECST
END_METHOD

METHOD CALL_S123_SELECTMODECSP
END_METHOD

METHOD CALL_S996_STOP
END_METHOD

METHOD CALL_S998_SERVICE
END_METHOD

METHOD CALL_S999_ERROR
END_METHOD

METHOD CALL_T002_READY
END_METHOD

METHOD CALL_T020_SYNCLINEVEL
END_METHOD

(* ---- _TM_WINDERDANCERCTRLBASE.fb ---- *)
FUNCTION_BLOCK _TM_WINDERDANCERCTRLBASE EXTENDS _TM_Winder
VAR_OUTPUT
	PPAR : POINTER TO _scPar_TM_WinderDancerCtrlHigh;
	PSF : POINTER TO _scSF_TM_WinderDancerCtrlHigh;
	PAP : POINTER TO _scAP_TM_WinderDancerCtrlHigh;
END_VAR
VAR_IN_OUT
	LRSETLINEVELDIAMCALC : LREAL;
	XTEACHUPPERPOS : BOOL;
	XTEACHLOWERPOS : BOOL;
	XDANCERCTRL : BOOL;
	XRESETICTRL : BOOL;
	LRACTDANCERPOSIN : LREAL;
	LRSETDANCERPOSSCALED : LREAL;
	LRDANCERPOSINFLUENCESCALED : LREAL;
	XDANCERREACHEDSETPOS : BOOL;
	XDANCERMAXPOS : BOOL;
	XDANCERMINPOS : BOOL;
	LRACTDANCERPOSSCALED : LREAL;
	LRSETDANCERPOSCTRLSCALEDOUT : LREAL;
	LRSETTENSCURVEOUT : LREAL;
END_VAR
VAR
	XRESETICTRL_INT : BOOL;
	XTEACHUPPERPOS_INT : BOOL;
	XTEACHLOWERPOS_INT : BOOL;
	XRESETTEACHDANCERPOS_INT : BOOL;
	XDANCERCTRL_INT : BOOL;
	LRSETDANCERPOSSCALED_INT : LREAL;
	LRDANCERPOSINFLUENCESCALED_INT : LREAL := 0.1;
	XTEACHDANCERLIMITS_OLD : BOOL;
	XTEACHUPPERPOS_INT_OLD : BOOL;
	XTEACHLOWERPOS_INT_OLD : BOOL;
	XRESETICTRL_OLD : BOOL;
	LRDANCERPOSCTRLRESETTIME_STORE : LREAL;
	LRDEVIATION_STORE : LREAL;
	SCPAR_INT : _scPar_TM_WinderDancerCtrlHigh;
	XDANCERCONTROLACTIVE_INT : BOOL;
	LRSETREELSPEEDFRWCTRL : LREAL;
	LRSETREELSPEEDDEVIATION : LREAL;
	LRDANCERPOSCTRLOUTVEL : LREAL;
	LRSETSPEEDTOTAL : LREAL;
	LRDANCERPOSREF : LREAL;
	LRDANCERPOSSCALED0TO1 : LREAL;
	LRFILTACTDANCERPOS : LREAL;
	LRFILTACTDANCERPOSSCALED : LREAL;
	LRACTDANCERVEL : LREAL;
	LRACTDANCERLINEVELCOMP : LREAL;
	XWARNING_DANCERLIMITSNOTTEACHED : BOOL;
	L_MB1P_RAMPGENERATORRESETICTRL : L_MC1P_RampGenerator;
	L_MB1P_DIFFERENTIATE1 : L_MC2P_Differentiate;
	L_MB1P_PROCESSCONTROLLER1 : L_CT1P_ProcessController;
	L_D94A_FILTERDANCERPOSIN : L_USPP_PT1Filter;
	L_D94A_FILTERLINEVELCOMP : L_USPP_PT1Filter;
	LRDANCERUPPERLIMIT_INT : LREAL;
	LRDANCERLOWERLIMIT_INT : LREAL;
	XUPPERPOSTEACHED : BOOL;
	XLOWERPOSTEACHED : BOOL;
	LRTEACHEDDANCERUPPERLIMIT_INT : LREAL;
	LRTEACHEDDANCERLOWERLIMIT_INT : LREAL;
END_VAR
END_FUNCTION_BLOCK

METHOD CALL_ALLOCPOINTADR
END_METHOD

METHOD CALL_CTRLREQACTIVE : BOOL
END_METHOD

METHOD CALL_ERRORHANDLER
END_METHOD

METHOD CALL_FBMETHODS
END_METHOD

METHOD CALL_FBMETHODS_WND
END_METHOD

METHOD CALL_FB_PROCESSCONTROLLER
END_METHOD

METHOD CALL_FB_PROCESSCONTROLLER_INPUT
END_METHOD

METHOD CALL_FB_RAMPGENERATOR_INPUT
END_METHOD

METHOD CALL_FB_WNDCALCDIAMETER_HOLDDIAMETER
END_METHOD

METHOD CALL_FB_WNDCALCDIAMETER_INPUT
END_METHOD

METHOD CALL_FILTERDANCERPOSIN
END_METHOD

METHOD CALL_FILTERLINEVELCOMP
END_METHOD

METHOD CALL_FIRSTCYCLE
END_METHOD

METHOD CALL_INITROUTINE
END_METHOD

METHOD CALL_INTERNALCTRL
END_METHOD

METHOD CALL_INTERNALCTRLNOTACTIVE
END_METHOD

METHOD CALL_OUTPUT
END_METHOD

METHOD CALL_OUTPUT_SF
END_METHOD

METHOD CALL_RAMPGENERATORRESETICTRL
END_METHOD

METHOD CALL_REQUESTS_EXT
END_METHOD

METHOD CALL_RESETCOMMANDS
END_METHOD

METHOD CALL_RESETOUTPUT
END_METHOD

METHOD CALL_RESETWARNINGS
END_METHOD

METHOD CALL_SDDIFFERENTIATE : BOOL
END_METHOD

METHOD CALL_SETSPEEDPOINT
END_METHOD

METHOD CALL_STATEMACHINE
END_METHOD

METHOD CALL_TEACHDANCER
END_METHOD

METHOD CALL_WNDTENSIONCURVE_INPUT
END_METHOD

METHOD GET_LRACTDANCERCTRLOUT : LREAL
END_METHOD

METHOD GET_LRACTDANCERLINEVELCOMP : LREAL
END_METHOD

METHOD GET_LRACTDANCERVEL : LREAL
END_METHOD

METHOD GET_LRSPEEDFORWARDCTRL : LREAL
END_METHOD

METHOD GET_LRSPEEDSETPOINT : LREAL
END_METHOD

METHOD GET_LRVELSETPOINT : LREAL
END_METHOD

METHOD GET_XLOWERPOSTEACHED : BOOL
VAR_OUTPUT
	LRTEACHPOSLOWERLIMIT : LREAL;
END_VAR
END_METHOD

METHOD GET_XUPPERPOSTEACHED : BOOL
VAR_OUTPUT
	LRTEACHPOSUPPERLIMIT : LREAL;
END_VAR
END_METHOD

METHOD CALL_RESTDANCERTEACHPOS
END_METHOD

METHOD LOAD_LRDANCERLOWERLIMIT
VAR_INPUT
	LRIN : LREAL := 0;
END_VAR
END_METHOD

METHOD LOAD_LRDANCERUPPERLIMIT
VAR_INPUT
	LRIN : LREAL := 0;
END_VAR
END_METHOD

METHOD SET_ALRPROCESSCTRLXVALUES
VAR_INPUT
	ALRPROCESSCTRLXVALUES : ARRAY [1..5] OF LREAL := [5(0)];
END_VAR
END_METHOD

METHOD SET_ALRPROCESSCTRLYVALUES
VAR_INPUT
	ALRPROCESSCTRLYVALUES : ARRAY [1..5] OF LREAL := [1, 4(0)];
END_VAR
END_METHOD

METHOD SET_LRPICTRLINTVALUE
VAR_INPUT
	LRIN : LREAL := 0;
END_VAR
END_METHOD

METHOD SET_LRPROCESSCTRLACC
VAR_INPUT
	LRPROCESSCTRLACC : LREAL := 0.0;
END_VAR
END_METHOD

METHOD SET_LRPROCESSCTRLDEC
VAR_INPUT
	LRPROCESSCTRLDEC : LREAL := 0.0;
END_VAR
END_METHOD

METHOD SET_LRPROCESSCTRLGAINADAPT
VAR_INPUT
	LRPROCESSCTRLGAINADAPT : LREAL := 1;
END_VAR
END_METHOD

METHOD SET_LRPROCESSCTRLINTVALUE
VAR_INPUT
	LRPROCESSCTRLINTVALUE : LREAL := 0.0;
END_VAR
END_METHOD

METHOD SET_LRPROCESSCTRLREDGAIN
VAR_INPUT
	LRPROCESSCTRLREDGAIN : LREAL := 0.0;
END_VAR
END_METHOD

METHOD SET_LRPROCESSCTRLREDRANGE
VAR_INPUT
	LRPROCESSCTRLREDRANGE : LREAL := 0.0;
END_VAR
END_METHOD

METHOD SET_RPROCESSCTRLDELAYTIME
VAR_INPUT
	RPROCESSCTRLDELAYTIME : REAL := 0.0;
END_VAR
END_METHOD

METHOD SET_RPROCESSCTRLRATEDTIME
VAR_INPUT
	RPROCESSCTRLRATEDTIME : REAL := 0.0;
END_VAR
END_METHOD

METHOD SET_XPICTRLLOADINTVALUE
VAR_INPUT
	XIN : BOOL := FALSE;
END_VAR
END_METHOD

METHOD SET_XPROCESSCTRLLOADINTVALUE
VAR_INPUT
	XPROCESSCTRLLOADINTVALUE : BOOL := FALSE;
END_VAR
END_METHOD

METHOD CALL_S000_CYCLIC
END_METHOD

METHOD CALL_S002_READY
END_METHOD

METHOD CALL_S020_SYNCLINEVEL
END_METHOD

METHOD CALL_S050_DANCERTRL
END_METHOD

METHOD CALL_S999_ERROR
END_METHOD

METHOD CALL_T002_READY
END_METHOD

METHOD CALL_T020_SYNCLINEVEL
END_METHOD

METHOD CALL_T050_DANCERTRL
END_METHOD

(* ---- _TM_WINDERDANCERCTRLHIGH.fb ---- *)
FUNCTION_BLOCK _TM_WINDERDANCERCTRLHIGH EXTENDS _TM_WinderDancerCtrlState
VAR_IN_OUT
	XEXECUTEIDENTMINERTIA : BOOL;
	XEXECUTEIDENTDIAM : BOOL;
	XADAPTSPDCTRLGAIN : BOOL;
	LRADAPTSPDCTRLGAINFACTOR : LREAL;
	LRIDENTMINERTIA : LREAL;
	LRSETSPDCTRLGAINADAPTOUT : LREAL;
END_VAR
VAR
	XEXECUTEIDENTMINERTIA_INT : BOOL;
	XEXECUTEIDENTDIAM_INT : BOOL;
	XADAPTSPDCTRLGAIN_INT : BOOL;
	LRADAPTSPDCTRLGAINFACTOR_INT : LREAL;
	WSTEPPER_DANCERCTRLSTOPMODE : WORD;
	LRTIME : LREAL;
	LRDIST : LREAL;
	LRDISTTOTARGET : LREAL;
	LRRELDIST : LREAL;
	LRSTOREACTPOS : LREAL;
	LRSETPOS_DIST_INT : LREAL;
	LRTARGETPOSITION : LREAL;
	LRVEL_INT : LREAL;
	LRACTFOLLOWINGERROR : LREAL;
	XDONEFROMIDENTMINERTIA : BOOL;
	XIDENTDIAM_LOADDIAM : BOOL;
	LRIDENTDIAM_SETDIAMETER : LREAL;
	EDANCERCTRLSTOPMODE_OLD : L_TT1P_DancerCtrlStopMode;
	XERROR_IDENTDIAMMAXDANCERPOS : BOOL;
	XERROR_ACTDANPOSBIGGERMAXDANPOS : BOOL;
	XERRORFOLLOWINGERRORSWITCHTOPOSCTRLDRIVE : BOOL;
	XERROR_IDENTIFICATIONDIAMETERFAILED : BOOL;
	XERROR_INVALIDDANCERMATERIALLENGTH : BOOL;
	XWARNING_INVALIDDANCERMATERIALLENGTH : BOOL;
	XWARNING_IDENTIFICATIONDIAMETERFAILED : BOOL;
	XWARNING_INVALIDLOADDIAM : BOOL;
	XWARNING_INVALIDIDENTMAXDANCERPOS : BOOL;
	XWARNING_ACTDANCERPOSBIGGERMAXDANCERPOS : BOOL;
	WIDENTDIAMCALCCYCLES : WORD;
	XIDENTMINERTIASPEELIMITS : BOOL;
	L_MB1P_IDENTMINERTIA1 : L_TB1P_IdentMInertia;
	L_MB1P_CURVESPEEDCTRLGAIN : L_USPP_Curve;
	FB_WINDERIDENTDIAMETER : L_MB1P_WinderIdentDiameter;
	FB_SETSPEEDCTRLADAPTVAL1 : L_MC1P_SetSpeedCtrlAdaptValue;
END_VAR
END_FUNCTION_BLOCK

METHOD CALL_CTRLREQACTIVE : BOOL
END_METHOD

METHOD CALL_ERRORHANDLER
END_METHOD

METHOD CALL_FBMETHODS_WND
END_METHOD

METHOD CALL_FB_CURVESPEEDCTRLGAIN
END_METHOD

METHOD CALL_FB_CURVESPEEDCTRLGAIN_INPUT
END_METHOD

METHOD CALL_FB_PROCESSCONTROLLER_INPUT
END_METHOD

METHOD CALL_FB_SETSPEEDCTRLADAPTVALUE
END_METHOD

METHOD CALL_FB_SETSPEEDCTRLADAPTVALUE_INPUT
END_METHOD

METHOD CALL_FB_WINDERIDENTDIAMETER
END_METHOD

METHOD CALL_FB_WINDERIDENTDIAMETER_INPUT
END_METHOD

METHOD CALL_FB_WNDCALCDIAMETER_INPUT
END_METHOD

METHOD CALL_FIRSTCYCLE
END_METHOD

METHOD CALL_INITROUTINE
END_METHOD

METHOD CALL_INTERNALCTRLACTIVE
END_METHOD

METHOD CALL_INTERNALCTRLNOTACTIVE
END_METHOD

METHOD CALL_LIMITEDINPUT
END_METHOD

METHOD CALL_OUTPUT
END_METHOD

METHOD CALL_REQUESTS_EXT
END_METHOD

METHOD CALL_RESETCOMMANDS
END_METHOD

METHOD CALL_RESETOUTPUT
END_METHOD

METHOD CALL_RESETWARNINGS
END_METHOD

METHOD CALL_SETSPEEDPOINT
END_METHOD

METHOD CALL_SETTORQUE
END_METHOD

METHOD CALL_STATEMACHINE
END_METHOD

METHOD CALL_WNDIDENTMINERTIA
END_METHOD

METHOD CALL_S000_CYCLIC
END_METHOD

METHOD CALL_S002_READY
END_METHOD

METHOD CALL_S014_MOVEABS
END_METHOD

METHOD CALL_S015_MOVEREL
END_METHOD

METHOD CALL_S040_IDENTMINERTIA
END_METHOD

METHOD CALL_S050_DANCERTRL
END_METHOD

METHOD CALL_S081_IDENTDIAMETER
END_METHOD

METHOD CALL_S996_STOP
END_METHOD

METHOD CALL_S999_ERROR
END_METHOD

METHOD CALL_T002_READY
END_METHOD

METHOD CALL_T050_DANCERTRL
END_METHOD

(* ---- _TM_WINDERDANCERCTRLSTATE.fb ---- *)
FUNCTION_BLOCK _TM_WINDERDANCERCTRLSTATE EXTENDS _TM_WinderDancerCtrlBase
VAR_IN_OUT
	XACCCMPS : BOOL;
	LRMINERTIAADAPT : LREAL;
	LRSETMINERTIAOUT : LREAL;
	LRSETACCTRQSCALEDOUT : LREAL;
END_VAR
VAR
	XACCCMPS_INT : BOOL;
	LRMINERTIAADAPT_INT : LREAL := 1;
	XDECOUPLINGACCCOMP : BOOL;
	LRSETACCTORQUE : LREAL;
	LRACTACCTORQUE : LREAL;
	XACCCMPSACTIVE_INT : BOOL;
	L_MB1P_ACCCOMP1 : L_TB1P_AccComp;
END_VAR
END_FUNCTION_BLOCK

METHOD CALL_FBMETHODS_WND
END_METHOD

METHOD CALL_FB_ACCCOMP : LREAL
END_METHOD

METHOD CALL_FB_ACCCOMP_INPUT : LREAL
END_METHOD

METHOD CALL_FIRSTCYCLE
END_METHOD

METHOD CALL_INTERNALCTRLNOTACTIVE
END_METHOD

METHOD CALL_OUTPUT
END_METHOD

METHOD CALL_OUTPUT_SF
END_METHOD

METHOD CALL_RESETCOMMANDS
END_METHOD

METHOD CALL_RESETOUTPUT
END_METHOD

METHOD CALL_SETTORQUE
END_METHOD

METHOD CALL_WNDTENSIONCURVE_INPUT
END_METHOD

METHOD GET_LRACTACCTRQ : LREAL
END_METHOD

METHOD CALL_S000_CYCLIC
END_METHOD

METHOD CALL_S010_JOGGING
END_METHOD

METHOD CALL_S020_SYNCLINEVEL
END_METHOD

(* ---- _TM_WINDERTENSIONCTRLBASE.fb ---- *)
FUNCTION_BLOCK _TM_WINDERTENSIONCTRLBASE EXTENDS _TM_Winder
VAR_OUTPUT
	PPAR : POINTER TO _scPar_TM_WinderTensionCtrlHigh;
	PSF : POINTER TO _scSF_TM_WinderTensionCtrlHigh;
	PAP : POINTER TO _scAP_TM_WinderTensionCtrlHigh;
END_VAR
VAR_IN_OUT
	XWINDINGDIRECTIONSTANDSTILL : BOOL;
	XTENSCTRL : BOOL;
	XFRICCMPS : BOOL;
	XACCCMPS : BOOL;
	LRMINERTIAADAPT : LREAL;
	XWNDSPDLIMIT : BOOL;
	LRSETMINERTIAOUT : LREAL;
	LRSETTENSSCALEDOUT : LREAL;
	LRSETTENSTRQSCALEDOUT : LREAL;
	LRSETFRICTRQSCALEDOUT : LREAL;
	LRSETACCTRQSCALEDOUT : LREAL;
END_VAR
VAR
	XTENSCTRL_INT : BOOL;
	XACCCMPS_INT : BOOL;
	XFRICCMPS_INT : BOOL;
	LRMINERTIAADAPT_INT : LREAL := 1;
	LRACTTENSIN_INT : LREAL := 0;
	LRFILTACTTENSIN : LREAL;
	XPICONTROLACTIVE_INT : BOOL;
	SCPAR_INT : _scPar_TM_WinderTensionCtrlHigh;
	WTENSRAMPLOADSTARTVALUEMODE : WORD;
	LRSETTENSSCALED : LREAL;
	LRPROCESSCTRLREDOUT : LREAL;
	LRSETPOINTTENSION : LREAL;
	LRSETTENSIONTORQUE : LREAL;
	LRSETFRICTIONTORQUE : LREAL;
	LRACTFRICTIONTORQUE : LREAL;
	LRSETACCTORQUE : LREAL;
	LRACTACCTORQUE : LREAL;
	LRSETLINEVELOFFSET : LREAL;
	LRSETTRQPOINT : LREAL;
	LRCALCWNDSPEEDUPPERLIMIT : LREAL;
	LRCALCWNDSPEEDLOWERLIMIT : LREAL;
	XACCCMPSACTIVE_INT : BOOL;
	XDECOUPLINGACCCOMP : BOOL;
	XDECOUPLINGFRICTIONCOMP : BOOL;
	XDECOUPLINGTENSION : BOOL;
	XWNDSPDLIMIT_OLD : BOOL;
	ICNTSPDLIMIT : INT;
	ISPDHYST : INT := 3;
	L_MB1P_ACCCOMP1 : L_TB1P_AccComp;
	L_D94A_FILTERREELSPEED : L_USPP_PT1Filter;
	L_D94A_FILTERREELSPEEDFRICTIONCOMP : L_USPP_PT1Filter;
END_VAR
END_FUNCTION_BLOCK

METHOD CALL_ALLOCPOINTADR
END_METHOD

METHOD CALL_CTRLREQACTIVE : BOOL
END_METHOD

METHOD CALL_FBMETHODS_WND
END_METHOD

METHOD CALL_FB_ACCCOMP : LREAL
END_METHOD

METHOD CALL_FB_ACCCOMP_INPUT : LREAL
END_METHOD

METHOD CALL_FB_RAMPGENERATOR_INPUT
END_METHOD

METHOD CALL_FB_WNDCALCDIAMETER_INPUT
END_METHOD

METHOD CALL_FILTERREELSPEED
END_METHOD

METHOD CALL_FIRSTCYCLE
END_METHOD

METHOD CALL_INTERNALCTRLNOTACTIVE
END_METHOD

METHOD CALL_OUTPUT
END_METHOD

METHOD CALL_OUTPUT_SF
END_METHOD

METHOD CALL_REQUESTS_EXT
END_METHOD

METHOD CALL_RESETCOMMANDS
END_METHOD

METHOD CALL_RESETOUTPUT
END_METHOD

METHOD CALL_SDRAMPGENERATOR_INPUT
END_METHOD

METHOD CALL_SETTORQUE
END_METHOD

METHOD CALL_SPEEDLIMIT
END_METHOD

METHOD CALL_STATEMACHINE
END_METHOD

METHOD CALL_WNDFRICTIONCOMPENSATION
END_METHOD

METHOD CALL_WNDTENSIONCURVE_INPUT
END_METHOD

METHOD GET_LRACTACCTRQ : LREAL
END_METHOD

METHOD GET_LRACTFRICTRQ : LREAL
END_METHOD

METHOD GET_LRACTTENSTRQ : LREAL
END_METHOD

METHOD GET_LRRAMPGENOUT : LREAL
END_METHOD

METHOD GET_LRSPEEDLOWERLIMIT : LREAL
END_METHOD

METHOD GET_LRSPEEDUPPERLIMIT : LREAL
END_METHOD

METHOD GET_LRTENSCTRLOUT : LREAL
END_METHOD

METHOD GET_LRTENSCURVEOUT : LREAL
END_METHOD

METHOD CALL_S000_CYCLIC
END_METHOD

METHOD CALL_S002_READY
END_METHOD

METHOD CALL_S010_JOGGING
END_METHOD

METHOD CALL_S020_SYNCLINEVEL
END_METHOD

METHOD CALL_S050_1_WNDFRICTIONCOMPENSATION
END_METHOD

METHOD CALL_S050_TENSIONCTRL
END_METHOD

METHOD CALL_T002_READY
END_METHOD

METHOD CALL_T020_SYNCLINEVEL
END_METHOD

METHOD CALL_T050_TENSIONCTRL
END_METHOD

(* ---- _TM_WINDERTENSIONCTRLHIGH.fb ---- *)
FUNCTION_BLOCK _TM_WINDERTENSIONCTRLHIGH EXTENDS _TM_WinderTensionCtrlState
VAR_IN_OUT
	XEXECUTEIDENTMINERTIA : BOOL;
	XADAPTSPDCTRLGAIN : BOOL;
	LRADAPTSPDCTRLGAINFACTOR : LREAL;
	LRIDENTMINERTIA : LREAL;
	LRSETSPDCTRLGAINADAPTOUT : LREAL;
END_VAR
VAR
	XEXECUTEIDENTMINERTIA_INT : BOOL;
	XADAPTSPDCTRLGAIN_INT : BOOL;
	LRADAPTSPDCTRLGAINFACTOR_INT : LREAL;
	WSTEPPER_TENSCTRLSTOPMODE : WORD;
	LRRELDIST : LREAL;
	LRSTOREACTPOS : LREAL;
	LRDISTTOTARGET : LREAL;
	LRACTFOLLOWINGERROR : LREAL;
	LRSETPOS_DIST_INT : LREAL;
	LRVEL_INT : LREAL;
	LRTARGETPOSITION : LREAL;
	LRDIST : LREAL;
	LRTIME : LREAL;
	LRSETVELOCITY_OLD : LREAL;
	XERRORFOLLOWINGERRORSWITCHTOPOSCTRLDRIVE : BOOL;
	ESTOPMODE_OLD : WORD;
	XIDENTMINERTIASPEELIMITS : BOOL;
	XDONEFROMIDENTMINERTIA : BOOL;
	L_MB1P_IDENTMINERTIA1 : L_TB1P_IdentMInertia;
	L_MB1P_CURVESPEEDCTRLGAIN : L_USPP_Curve;
	FB_SETSPEEDCTRLADAPTVAL1 : L_MC1P_SetSpeedCtrlAdaptValue;
END_VAR
END_FUNCTION_BLOCK

METHOD CALL_CTRLREQACTIVE : BOOL
END_METHOD

METHOD CALL_ERRORHANDLER
END_METHOD

METHOD CALL_FBMETHODS_WND
END_METHOD

METHOD CALL_FB_CURVESPEEDCTRLGAIN
END_METHOD

METHOD CALL_FB_CURVESPEEDCTRLGAIN_INPUT
END_METHOD

METHOD CALL_FB_SETSPEEDCTRLADAPTVALUE
END_METHOD

METHOD CALL_FB_SETSPEEDCTRLADAPTVALUE_INPUT
END_METHOD

METHOD CALL_FIRSTCYCLE
END_METHOD

METHOD CALL_INITROUTINE
END_METHOD

METHOD CALL_INTERNALCTRLNOTACTIVE
END_METHOD

METHOD CALL_LIMITEDINPUT
END_METHOD

METHOD CALL_OUTPUT
END_METHOD

METHOD CALL_REQUESTS_EXT
END_METHOD

METHOD CALL_RESETCOMMANDS
END_METHOD

METHOD CALL_RESETOUTPUT
END_METHOD

METHOD CALL_SETTORQUE
END_METHOD

METHOD CALL_STATEMACHINE
END_METHOD

METHOD CALL_WNDIDENTMINERTIA
END_METHOD

METHOD CALL_S000_CYCLIC
END_METHOD

METHOD CALL_S002_READY
END_METHOD

METHOD CALL_S014_MOVEABS
END_METHOD

METHOD CALL_S015_MOVEREL
END_METHOD

METHOD CALL_S040_IDENTMINERTIA
END_METHOD

METHOD CALL_S050_TENSIONCTRL
END_METHOD

METHOD CALL_S996_STOP
END_METHOD

METHOD CALL_S999_ERROR
END_METHOD

METHOD CALL_T002_READY
END_METHOD

METHOD CALL_T050_TENSIONCTRL
END_METHOD

(* ---- _TM_WINDERTENSIONCTRLSTATE.fb ---- *)
FUNCTION_BLOCK _TM_WINDERTENSIONCTRLSTATE EXTENDS _TM_WinderTensionCtrlBase
VAR_IN_OUT
	ALRFRICTIONCURVE1 : ARRAY [1..66] OF LREAL;
	ALRFRICTIONCURVE2 : ARRAY [1..66] OF LREAL;
	ALRFRICTIONCURVE3 : ARRAY [1..66] OF LREAL;
	ALRFRICTIONCURVE4 : ARRAY [1..66] OF LREAL;
	XRESETPICTRL : BOOL;
	XRESETICTRL : BOOL;
	LRACTTENSIN : LREAL := 0;
	LRSETFRICADAPT : LREAL;
	LRTENSCTRLINFLUENCE : LREAL := 0;
	XEXECUTEIDENTFRIC : BOOL;
	LRACTTENSSCALED : LREAL := 0;
	LRSETTENSCTRLSCALEDOUT : LREAL;
END_VAR
VAR
	XRESETPICTRL_INT : BOOL;
	XRESETPICTRL_OLD : BOOL;
	XRESETICTRL_INT : BOOL;
	XRESETICTRL_OLD : BOOL;
	LRTENSCTRLRESETTIME_STORE : LREAL;
	LRDEVIATION_STORE : LREAL;
	XEXECUTEIDENTFRIC_INT : BOOL;
	LRTENSCTRLINFLUENCE_INT : LREAL := 0;
	LRSETFRICADAPT_INT : LREAL;
	LRTENSPICTRLOUT : LREAL;
	XPIDENABLE_INT : BOOL;
	XPIDRESET_INT : BOOL;
	XPIDLOADACTVLAUE_INT : BOOL;
	XPIDLRESETICTRLACTIVE_INT : BOOL;
	XPIDLRESETPICTRLACTIVE_INT : BOOL;
	L_MB1P_RAMPGENERATORRESETICTRL : L_MC1P_RampGenerator;
	L_MB1P_RAMPGENERATORRESETPICTRL : L_MC1P_RampGenerator;
	XRAMPGENSETVALUEFORPICTRLACTIVE : BOOL;
	WRESETPICTRL_STEPPER : WORD;
	L_MB1P_PROCESSCONTROLLER1 : L_CT1P_ProcessController;
	L_MB1P_FRICTIONCOMPENSATION1 : L_TB1P_FrictionCompensation;
	L_D94A_FILTERTENSIN : L_USPP_PT1Filter;
END_VAR
END_FUNCTION_BLOCK

METHOD CALL_CTRLREQACTIVE : BOOL
END_METHOD

METHOD CALL_ERRORHANDLER
END_METHOD

METHOD CALL_FBMETHODS_WND
END_METHOD

METHOD CALL_FB_PROCESSCONTROLLER
END_METHOD

METHOD CALL_FB_PROCESSCONTROLLER_INPUT
END_METHOD

METHOD CALL_FB_RAMGENERATORRESETPICTRL
END_METHOD

METHOD CALL_FB_RAMPGENERATORRESETICTRL
END_METHOD

METHOD CALL_FB_RAMPGENERATORRESETICTRL_INPUT
END_METHOD

METHOD CALL_FB_RAMPGENERATORRESETPICTRL_INPUT
END_METHOD

METHOD CALL_FILTERTENSIN
END_METHOD

METHOD CALL_FIRSTCYCLE
END_METHOD

METHOD CALL_INTERNALCTRL
END_METHOD

METHOD CALL_INTERNALCTRLNOTACTIVE
END_METHOD

METHOD CALL_OUTPUT
END_METHOD

METHOD CALL_OUTPUT_SF
END_METHOD

METHOD CALL_REQUESTS_EXT
END_METHOD

METHOD CALL_RESETCOMMANDS
END_METHOD

METHOD CALL_RESETOUTPUT
END_METHOD

METHOD CALL_SETSPEEDPOINT
END_METHOD

METHOD CALL_STATEMACHINE
END_METHOD

METHOD CALL_WNDFRICTIONCOMPENSATION
END_METHOD

METHOD CALL_WNDTENSIONCURVE_INPUT
END_METHOD

METHOD SET_ALRPROCESSCTRLXVALUES
VAR_INPUT
	ALRPROCESSCTRLXVALUES : ARRAY [1..5] OF LREAL := [5(0)];
END_VAR
END_METHOD

METHOD SET_ALRPROCESSCTRLYVALUES
VAR_INPUT
	ALRPROCESSCTRLYVALUES : ARRAY [1..5] OF LREAL := [1, 4(0)];
END_VAR
END_METHOD

METHOD SET_LRPICTRLINTVALUE
VAR_INPUT
	LRIN : LREAL := 0;
END_VAR
END_METHOD

METHOD SET_LRPROCESSCTRLACC
VAR_INPUT
	LRPROCESSCTRLACC : LREAL := 0.0;
END_VAR
END_METHOD

METHOD SET_LRPROCESSCTRLDEC
VAR_INPUT
	LRPROCESSCTRLDEC : LREAL := 0.0;
END_VAR
END_METHOD

METHOD SET_LRPROCESSCTRLGAINADAPT
VAR_INPUT
	LRPROCESSCTRLGAINADAPT : LREAL := 1;
END_VAR
END_METHOD

METHOD SET_LRPROCESSCTRLINTVALUE
VAR_INPUT
	LRPROCESSCTRLINTVALUE : LREAL := 0.0;
END_VAR
END_METHOD

METHOD SET_LRPROCESSCTRLREDGAIN
VAR_INPUT
	LRPROCESSCTRLREDGAIN : LREAL := 0.0;
END_VAR
END_METHOD

METHOD SET_LRPROCESSCTRLREDRANGE
VAR_INPUT
	LRPROCESSCTRLREDRANGE : LREAL := 0.0;
END_VAR
END_METHOD

METHOD SET_RPROCESSCTRLDELAYTIME
VAR_INPUT
	RPROCESSCTRLDELAYTIME : REAL := 0.0;
END_VAR
END_METHOD

METHOD SET_RPROCESSCTRLRATEDTIME
VAR_INPUT
	RPROCESSCTRLRATEDTIME : REAL := 0.0;
END_VAR
END_METHOD

METHOD SET_XPICTRLLOADINTVALUE
VAR_INPUT
	XIN : BOOL := FALSE;
END_VAR
END_METHOD

METHOD SET_XPROCESSCTRLLOADINTVALUE
VAR_INPUT
	XPROCESSCTRLLOADINTVALUE : BOOL := FALSE;
END_VAR
END_METHOD

METHOD CALL_S000_CYCLIC
END_METHOD

METHOD CALL_S002_READY
END_METHOD

METHOD CALL_S030_IDENTFRICTION
END_METHOD

METHOD CALL_S050_1_WNDFRICTIONCOMPENSATION
END_METHOD

METHOD CALL_S050_TENSIONCTRL
END_METHOD

METHOD CALL_S999_ERROR
END_METHOD

METHOD CALL_T002_READY
END_METHOD

METHOD CALL_T020_SYNCLINEVEL
END_METHOD

(* ---- GLOBALTEXTLIST.fb ---- *)
FUNCTION_BLOCK GLOBALTEXTLIST
VAR
	M_TEXTLISTFILE : STRING(255);
	_STNAMESPACE : STRING;
END_VAR
END_FUNCTION_BLOCK

(* ---- L_MB1P_CALCOSCILATIONCOMPPARAMETER.fb ---- *)
FUNCTION_BLOCK L_MB1P_CALCOSCILATIONCOMPPARAMETER
VAR_INPUT
	XEXECUTE : BOOL;
	LRSETPOS : LREAL;
	LRSETLOAD : LREAL;
END_VAR
VAR_OUTPUT
	XBUSY : BOOL;
	XVALID : BOOL;
	XCALCPARAMACTIVE : BOOL;
	XDISABLEDOSCCOMPDATA : BOOL;
	LREIGENFREQUENCY : LREAL;
	LRAMPRATIO : LREAL;
END_VAR
VAR_IN_OUT
	ASCOSCCOMPDATA : ARRAY [1..8] OF L_TT1P_OscillationCompensationData;
END_VAR
VAR
	XEXECUTE_OLD : BOOL;
	WSTATE : WORD;
	XENTRY : BOOL;
	LRSETPOS_INT : LREAL;
	LRSETLOAD_INT : LREAL;
	INUMOFVALIDDATA : INT;
	AIPARAIDX : ARRAY [1..c_iMaxN, 1..c_iMaxN] OF INT;
	IDX1 : INT;
	IDX2 : INT;
	IDX3 : INT;
	IDX4 : INT;
	IDX_LINKS : INT;
	IDX_RECHTS : INT;
	IDX_OBEN : INT;
	IDX_UNTEN : INT;
	IN : INT;
	IM : INT;
	LRTOLERANZPOS : LREAL;
	IDX_LINKS_DATA : INT;
	IDX_RECHTS_DATA : INT;
	IDX_OBEN_DATA : INT;
	IDX_UNTEN_DATA : INT;
	LRPOSSCLAED_TMP : LREAL;
	LRLOADSCLAED_TMP : LREAL;
	LRPOS0 : LREAL;
	LRPOS1 : LREAL;
	LRDIFFPOS : LREAL;
	LRLOAD0 : LREAL;
	LRLOAD1 : LREAL;
	LRDIFFLOAD : LREAL;
	ALREIGENFREQ2D : ARRAY [1..2, 1..2] OF LREAL;
	ALRAMPRATION2D : ARRAY [1..2, 1..2] OF LREAL;
	C_IMAXN : INT := 8;
END_VAR
END_FUNCTION_BLOCK

(* ---- L_MB1P_CALCULATETPCOMPENSATIONFACTOR.fb ---- *)
FUNCTION_BLOCK L_MB1P_CALCULATETPCOMPENSATIONFACTOR
VAR_OUTPUT
	LRFACTOR : LREAL;
	LRCOMPENSATIONCYCLES : LREAL;
END_VAR
VAR_IN_OUT
	TPAXIS : Axis_Ref;
END_VAR
VAR
	LRSETPOSARRAY : ARRAY [0..15] OF LREAL;
	BYCOUNTER : BYTE;
	LRTEMP : LREAL;
	LRPOSDIFF : LREAL;
	LRSETACTDIFF : LREAL;
	XERRORINVALIDAXIS : BOOL;
	LRSETPOS : LREAL;
	LRACTPOS : LREAL;
	LRCYCLELENGTH : LREAL;
	LRADDITIONALCORRECTION : LREAL;
	LRTEMP2 : LREAL;
	XINCREMENTCYCLES : BOOL;
END_VAR
END_FUNCTION_BLOCK

METHOD SEARCHARRAY
END_METHOD

(* ---- L_MB1P_CAMCREATOR.fb ---- *)
FUNCTION_BLOCK L_MB1P_CAMCREATOR
VAR_INPUT
	XENABLEINTERNALCAMTABLE : BOOL;
	XEXECUTE : BOOL;
	PCAMPOINTS : POINTER TO L_MC2P_CamDataXYVA;
	INUMOFPOINTS : INT;
	LRMASTERMAXVEL : LREAL;
	LRMASTERMAXACC : LREAL;
	LRMASTERSCALING : LREAL := 1;
	LRSLAVESCALING : LREAL := 1;
END_VAR
VAR_OUTPUT
	XINTERNALCAMTABLELACTIVE : BOOL;
	XERROR : BOOL;
	EERRORID : L_IE1P_Error;
	XBUSY : BOOL;
	XDONE : BOOL;
	CAMTABLEOUT : MC_CAM_REF;
	LRSLAVEMAXPOS : LREAL;
	LRSLAVEMINPOS : LREAL;
	LRSLAVEMAXVEL : LREAL;
	LRSLAVEMINVEL : LREAL;
	LRSLAVEMAXACC : LREAL;
	LRSLAVEMINACC : LREAL;
END_VAR
VAR_IN_OUT
	SLAVE : AXIS_REF;
END_VAR
VAR
	EFMSTATE : L_MB1P_States := L_MB1P_States.INIT;
	SMC_CAMBOUNDS1 : L_MC2P_BoundsCam;
	SMC_CAMBOUNDSINIT : L_MC2P_BoundsCam;
	CAMREF : L_MC2P_CamRefFromStruct;
	PCAMPOINTS_INT : POINTER TO L_MC2P_CamDataXYVA;
	INUMOFPOINTS_INT : INT;
	XINTERNALCONTROL : BOOL;
	XEXECUTE_OLD : BOOL;
	ASCCAMPOINTS : ARRAY [0..30] OF L_MC2P_CamDataXYVA;
	XINVALIDCAMTABLE : BOOL;
	XVISUACTIVE : BOOL := TRUE;
	DIFRAME : DINT;
	DIFRAME_OLD : DINT;
	ARVISPOINTLINES : ARRAY [1..10] OF L_MC2P_CamDataXYVA;
	IVISUTABLESETPOS : INT := 0;
	IVISUTABLESETPOS_OLD : INT := 0;
	IVISUTABLEMAXPOS : INT := 30;
	IVISSHOWLINESNO : INT;
	XVISPOINTMIN : BOOL;
	XVISPOINTMAX : BOOL;
	XVISUSETPOSUP : BOOL;
	XVISUSETPOSDOWN : BOOL;
	XVISUSETPOSUP_OLD : BOOL;
	XVISUSETPOSDOWN_OLD : BOOL;
	XSCROLBUTTENACTIVE : BOOL;
	TSETTIME : TIME := TIME#400ms;
	TON_SCROLBUTTEN : TON;
END_VAR
END_FUNCTION_BLOCK

METHOD CALL_CAMBOUNDS
VAR_IN_OUT
	SLAVE : AXIS_REF;
END_VAR
END_METHOD

METHOD CALL_CAMREF
END_METHOD

METHOD CALL_CAMTABLEEQUIDISTANT
END_METHOD

METHOD CALL_CAMTABLENONEQUIDISTANT
END_METHOD

METHOD CALL_CAMTABLEPOLYNOMIAL
END_METHOD

METHOD CALL_ERRORHANDLER
END_METHOD

METHOD CALL_FBMETHODS
VAR_IN_OUT
	SLAVE : AXIS_REF;
END_VAR
END_METHOD

METHOD CALL_INTERNALCTRL
END_METHOD

METHOD CALL_OUTPUT
END_METHOD

METHOD CALL_RESETCOMMANDS
VAR_IN_OUT
	SLAVE : AXIS_REF;
END_VAR
END_METHOD

METHOD CALL_RESETOUTPUT
END_METHOD

METHOD CALL_STATEMACHINE
END_METHOD

METHOD CALL_VIS_TON_SCROLBUTTEN
END_METHOD

METHOD CALL_VISUTABCTRL
END_METHOD

METHOD CALL_VISUUPDATETAB
END_METHOD

METHOD DISABALE_VISU
END_METHOD

METHOD ENABLE_VISU
END_METHOD

METHOD CALL_S000_CYCLIC
END_METHOD

METHOD CALL_S001_INIT
END_METHOD

METHOD CALL_S002_READY
END_METHOD

(* ---- L_MB1P_CAMTABLEINFO.fb ---- *)
FUNCTION_BLOCK L_MB1P_CAMTABLEINFO
VAR_INPUT
	XENABLE : BOOL;
	CAMTABLE : MC_CAM_REF;
	LRMASTERMAXVEL : LREAL := 100;
	LRMASTERMAXACC : LREAL := 1000;
	LRMASTERSCALING : LREAL := 1;
	LRSLAVESCALING : LREAL := 1;
END_VAR
VAR_OUTPUT
	XBUSY : BOOL;
	XDONE : BOOL;
	XCAMTABLEVALID : BOOL;
	LRMASTERSTARTPOS : LREAL;
	LRMASTERENDPOS : LREAL;
	LRSLAVESTARTPOS : LREAL;
	LRSLAVEENDPOS : LREAL;
	LRSLAVEMAXPOS : LREAL;
	LRSLAVEMINPOS : LREAL;
	LRSLAVEMAXVEL : LREAL;
	LRSLAVEMINVEL : LREAL;
	LRSLAVEMAXACC : LREAL;
	LRSLAVEMINACC : LREAL;
END_VAR
VAR_IN_OUT
	SLAVEAXIS : AXIS_REF;
END_VAR
VAR
	ESTATE : L_MB1P_States := L_MB1P_States.INIT;
	CAMTABLE_INT : MC_CAM_REF;
	PCAMDATA_INT : POINTER TO L_MC2P_CamData;
	LRMASTERMAXVEL_INT : LREAL := 0;
	LRMASTERMAXACC_INT : LREAL := 0;
	LRMASTERSCALING_INT : LREAL := 0;
	LRSLAVESCALING_INT : LREAL := 0;
	XENABLE_OLD : BOOL;
	SMC_CAMBOUNDS1 : L_MC2P_BoundsCam;
	XCALCNEWVALUES : BOOL;
END_VAR
END_FUNCTION_BLOCK

METHOD CALC_STARTENDVALUES
END_METHOD

METHOD CALL_CAMBOUNDS
END_METHOD

METHOD CALL_FBMETHODS
END_METHOD

METHOD CALL_OUTPUT
END_METHOD

METHOD CALL_RESETCOMMANDS
END_METHOD

METHOD CALL_RESETOUTPUT
END_METHOD

METHOD CALL_STATEMACHINE
END_METHOD

METHOD GET_XCALCNEWVALUES : BOOL
END_METHOD

METHOD GET_XCRITICALCYCLE : BOOL
END_METHOD

(* ---- L_MB1P_CHECKMODULOOVERRUN.fb ---- *)
FUNCTION_BLOCK L_MB1P_CHECKMODULOOVERRUN
VAR_INPUT
	LRSETPOS : LREAL;
	LRSETVEL : LREAL;
	LRPERIOD : LREAL;
END_VAR
VAR_OUTPUT
	XOVERRUNPOS : BOOL;
	XOVERRUNNEG : BOOL;
END_VAR
VAR
	ALRMEM : ARRAY [1..7] OF LREAL;
END_VAR
END_FUNCTION_BLOCK

METHOD CALL_CHECKMODULOOVERRUN
VAR_IN_OUT
	LRSETPOS : LREAL;
	LRSETVEL : LREAL;
	LRPERIOD : LREAL;
	XOVERRUNPOS : BOOL;
	XOVERRUNNEG : BOOL;
	ALRMEM : ARRAY [1..7] OF LREAL;
END_VAR
END_METHOD

(* ---- L_MB1P_CLUTCHEXTENDEDBASE.fb ---- *)
FUNCTION_BLOCK L_MB1P_CLUTCHEXTENDEDBASE EXTENDS L_MC2P_ClutchBasic
VAR_INPUT
	XENABLE : BOOL;
	XCLUTCHCLOSE : BOOL;
	XCLUTCHOPENINSTANT : BOOL;
	ECLUTCHMODE : L_MB1P_ClutchMode := L_MB1P_ClutchMode.ramp_pos;
	ECLUTCHDIRECTION : L_MC2P_ClutchDirection := L_MC2P_ClutchDirection.mcCurrentDirection;
	EDIRECTION : L_MB1P_Direction := 0;
	LRCYCMASTERPOS : LREAL;
	LRCYCMASTERVEL : LREAL;
	LRCYCMASTERACC : LREAL;
	LRCYCSLAVEPOS : LREAL;
	LRCYCSLAVEVEL : LREAL;
	LRCYCSLAVEACC : LREAL;
	LROPENINSTANTDEC : LREAL;
	LRMASTERCLOSEPOS : LREAL;
	LRMASTERCLOSEDIST : LREAL := 100;
	LRSLAVECLOSEDIST : LREAL := 100;
	LRMASTEROPENDIST : LREAL := 100;
	LRSLAVEOPENDIST : LREAL := 100;
	LRSLAVEOPENPOS : LREAL;
	LRCLOSETIME : LREAL := 5;
	LROPENTIME : LREAL := 5;
	LRCLUTCHVEL : LREAL := 100;
	LRCLUTCHACC : LREAL := 1000.0;
	LRCLUTCHDEC : LREAL := 1000.0;
	LRCLUTCHJERK : LREAL := 1000000.0;
	LRVELTOLERANCE : LREAL := 1;
	LRAXESCYCLELENGTH : LREAL := 360;
	EMASTERTRAVERSINGRANGE : L_MC1P_TraversingRange;
	LRCYCLETIME : LREAL := 0.001;
END_VAR
VAR_OUTPUT
	XERROR : BOOL;
	EERRORID : L_IE1P_Error;
	XBUSY : BOOL;
	XDONE : BOOL;
	XSYNCHRONISED : BOOL;
	XCLUTCHACTIVE : BOOL;
	LRSETSLAVEPOSOUT : LREAL;
	LRSETSLAVEVELOUT : LREAL;
	LRSETSLAVEACCOUT : LREAL;
	LRSETSLAVEOFFSETOUT : LREAL;
	LRX0 : LREAL;
	LRX1 : LREAL;
	LRY0 : LREAL;
	LRY1 : LREAL;
	LRX0N : LREAL;
	LRX1N : LREAL;
	LRY0N : LREAL;
	LRY1N : LREAL;
	LRX0P : LREAL;
	LRX1P : LREAL;
	LRY0P : LREAL;
	LRY1P : LREAL;
END_VAR
VAR
	EAXESTRAVERSINGRANGE_INT : L_MC1P_TraversingRange;
	ECLUTCHMODE_INT : L_MB1P_ClutchMode;
	ECLUTCHDIRECTION_INT : L_MB1P_ClutchDirection;
	LRSETSLAVEOFFSET_CLUTCHREL : LREAL;
	LRSETSLAVEOFFSET_INT : LREAL;
	LRSETMASTEROFFSET_OVERRUN : LREAL;
	LRCYCLETIME_INT : LREAL;
	XCLUTCHOPENINSTANT_ACTIVE : BOOL;
	LROPENINSTANTDEC_INT : LREAL;
	XCLUTCHBASICENABLE : BOOL;
	LRTEMP : LREAL;
	LRDELTASETENDPOS : LREAL;
	LRDELTASETENDPOS_OLD : LREAL;
	LRDELTASETENDPOS_OLD2 : LREAL;
	XCLUTCHMASTERVELPOSITIVE : BOOL;
	XMASTERREVERSING : BOOL;
	XCLUTCHBASIC_EXECUTE_OLD : BOOL;
	XCLUTCHCLOSE_OLD : BOOL;
	XCLUTCHOPENINSTANT_OLD : BOOL;
	XBUSY_OLD : BOOL;
	XENABLE_OLD : BOOL;
	LRCYCMASTERPOS_OLD : LREAL;
	LRMASTERVELADD : LREAL;
	LRMASTERVELADDSYNC : LREAL;
	LRSLAVESTARTPOS : LREAL;
	LRMASTERCLOSEPOS_INT : LREAL;
	LRMASTERCLOSEDIST_INT : LREAL;
	LRSLAVECLOSEDIST_INT : LREAL;
	LRSLAVEOPENDIST_INT : LREAL;
	LRSLAVEOPENPOS_INT : LREAL;
	XSYNCMODEIN_INT : BOOL;
	LRCLUTCHTIME : LREAL;
	XCLUTCHPOSMODE_INT : BOOL := TRUE;
	LRCLUTCHVEL_INT : LREAL := 100;
	LRCLUTCHACC_INT : LREAL := 1000.0;
	LRCLUTCHDEC_INT : LREAL := 1000.0;
	LRCLUTCHJERK_INT : LREAL := 1000000.0;
	EMASTERDIRECTION_INT : L_MC2P_ClutchDirection;
	IMASTERMOVEMENTTYPE_INT : INT;
	XREVERSEALLOWED_INT : BOOL;
	XPERIODIC_INT : BOOL;
	LRSLAVEJERK : LREAL;
	ESTATE : L_MB1P_States := L_MB1P_States.INIT;
	XSTATEENTRY : BOOL;
	XSETPARAGAIN : BOOL;
	XERROR_LOCK : BOOL;
	EERRORID_LOCK : L_IE1P_Error;
	LRTOLERANCE : LREAL;
	ICYCLECNTAFTEREXECUTE : INT;
	XRESTART_INT : BOOL;
	SCCYCMASTER : L_MC2P_AxisProfile;
	SCCYCSLAVE : L_MC2P_AxisProfile;
	SCSETSLAVEOUT : L_MC2P_AxisProfile;
	SCSETSLAVEOUT_OLD : L_MC2P_AxisProfile;
	PSCSETSLAVEOUT : POINTER TO L_MC2P_AxisProfile;
	EMASTERDIRECTION : L_MC2P_ClutchDirection;
	XCLUTCHBASIC_DONE : BOOL;
	XCLUTCHBASIC_WARNINGCANTPREVENTREVERSE : BOOL;
	XCLUTCHBASIC_ERROR : BOOL;
	ECLUTCHBASIC_ERRORIDCLUTCH : L_IE1P_Error;
	XCLUTCHBASIC_BUSY : BOOL;
	XCLUTCHBASIC_CLUTCHACTIVE : BOOL;
	XCLUTCHBASIC_PERIODIC : BOOL;
	XCLUTCHBASIC_REVERSEALLOWED : BOOL;
	ECLUTCHBASIC_MASTERAXISTYPE : L_MC1P_TraversingRange;
	XCLUTCHBASIC_EXECUTE : BOOL;
	FB_CHECKMODULOOVERRUN : L_MB1P_CheckModuloOverrun;
	XHALT_OLD : BOOL;
	XHALTBUSYINT : BOOL;
	XHALTDONEINT : BOOL;
	XSIMPLEFUNRAMPSLAVEDIST : BOOL := TRUE;
	LRSETSLAVEOFFSET_CLUTCHRELENTRY : LREAL;
	XRAMPDISTABSVIALINEAR : BOOL;
	XCLUTCHBASIC_BUSY_OLD : BOOL;
	XCLUTCHMASTERVELPOSITIVE_OLD : BOOL;
	XMASTERINSIDEXSIZE : BOOL;
	XMASTERINSIDEXSIZE_OLD : BOOL;
	XMASTERINSIDEXSIZEP : BOOL;
	XMASTERINSIDEXSIZEP_OLD : BOOL;
	XMASTERINSIDEXSIZEN : BOOL;
	XMASTERINSIDEXSIZEN_OLD : BOOL;
	XMASTERSTANDSTILL : BOOL;
	XCLUTCHDIRECTIONPOSITIVE : BOOL;
	ALRKOEF : ARRAY [0..5] OF LREAL;
	LRXFACTORN : LREAL;
	LRYFACTORN : LREAL;
	LRSETSLAVEOFFSET_CLUTCHRELN : LREAL;
	LRXFACTORP : LREAL;
	LRYFACTORP : LREAL;
	LRSETSLAVEOFFSET_CLUTCHRELP : LREAL;
	LRXFACTOR : LREAL;
	LRYFACTOR : LREAL;
	LRXSCALED : LREAL;
	LRYSCALED : LREAL;
	LRYSCALED_OLD : LREAL;
	LRYSCALEDDIFF : LREAL;
	LRSETYPOS : LREAL;
	LRSETYPOS_OLD : LREAL;
	LRSETYVEL : LREAL;
	LRSETYVEL_OLD : LREAL;
	LRSETYACC : LREAL;
	XCLUTCHDIRECTIONPOSITIVE_OLD : BOOL;
	LRMASTERCYCLELENGTH : LREAL;
	LRDUMMY : LREAL;
	LRCYCMASTERVEL_OLD : LREAL;
	WRAMPVELLACCSTEPPER : WORD;
	XNOREVERSEACTIVE : BOOL;
	XHALT_BUSY : BOOL;
	XHALT_DONE : BOOL;
	XSLAVEHALT : BOOL;
	C_ALRKOEF_SYNCIN : ARRAY [0..5] OF LREAL := [0, 0, 0, 1, -0.5, 0];
	C_ALRKOEF_SYNCOUT : ARRAY [0..5] OF LREAL := [0, 1, 0, -1, 0.5, 0];
END_VAR
END_FUNCTION_BLOCK

METHOD CALL_ALLOCPOINTADR
END_METHOD

METHOD CALL_CLUTCHCLOSEMODE
END_METHOD

METHOD CALL_CLUTCHOPENMODE
END_METHOD

METHOD CALL_ERRORHANDLER
END_METHOD

METHOD CALL_FBMETHODS
END_METHOD

METHOD CALL_FB_CHECKMODULOOVERRUN
END_METHOD

METHOD CALL_FB_CLUTCHBASIC
END_METHOD

METHOD CALL_FB_CLUTCHBASIC_INPUTSMASTER
END_METHOD

METHOD CALL_FB_CLUTCHBASIC_OPENINSTANT
END_METHOD

METHOD CALL_FB_CLUTCHBASIC_RAMPABS
END_METHOD

METHOD CALL_FB_CLUTCHBASIC_RAMPABS_TARGETPOS
END_METHOD

METHOD CALL_FB_CLUTCHBASIC_RAMPPOS
END_METHOD

METHOD CALL_FB_CLUTCHBASIC_RAMPREL
END_METHOD

METHOD CALL_FB_CLUTCHBASIC_RAMPSLAVEDIST
END_METHOD

METHOD CALL_FB_CLUTCHBASIC_RAMPTIME
END_METHOD

METHOD CALL_FB_CLUTCHBASIC_RAMPVELLACC
END_METHOD

METHOD CALL_FB_CLUTCHBASIC_RELATIVE
END_METHOD

METHOD CALL_MODULOTOLINEARMASTERPOS
END_METHOD

METHOD CALL_OUTPUT
END_METHOD

METHOD CALL_RAMPRELDIESTREL_CALCCOEFX0X1Y0Y1
END_METHOD

METHOD CALL_RAMPRELDISTABS_CALCCOEFX0X1Y0Y1
END_METHOD

METHOD CALL_RAMPRELDISTABS_CORRX0X1FORMODULOMASTER
END_METHOD

METHOD CALL_RAMPSLAVEDIST_ABS
END_METHOD

METHOD CALL_RAMPSLAVEDIST_REL
END_METHOD

METHOD CALL_RAMPSLAVEDIST_SETYPOSOUT
END_METHOD

METHOD CALL_RESETCLUTCH
END_METHOD

METHOD CALL_RESETCOMMANDS
END_METHOD

METHOD CALL_RESETOUTPUT
END_METHOD

METHOD CALL_SETCLUTCHCLOSEPAR
END_METHOD

METHOD CALL_SETCLUTCHCLOSEPAR_OLD
END_METHOD

METHOD CALL_SETCLUTCHOPENPAR
END_METHOD

METHOD CALL_SETCLUTCHOPENPAR_OLD
END_METHOD

METHOD CALL_STATEMASHINE
END_METHOD

METHOD SET_CLUTCHOFFSET : BOOL
VAR_INPUT
	LRIN : LREAL := 0;
END_VAR
END_METHOD

METHOD SLAVEHALT
VAR_INPUT
	XHALT : BOOL;
	SCACTSLAVE : L_MC2P_AxisProfile;
	LRMAXVELDIFF : LREAL;
	LRMAXACC : LREAL;
	LRMAXDEC : LREAL;
	LRJERK : LREAL;
	LRCYCLETIME : LREAL;
END_VAR
VAR_OUTPUT
	SCOUTPUTSLAVE : L_MC2P_AxisProfile;
	XBUSY : BOOL;
	XDONE : BOOL;
	XERROR : BOOL;
	EERRORID : L_IE1P_Error;
END_VAR
END_METHOD

METHOD CALL_S000_CYCLIC
END_METHOD

METHOD CALL_S001_INIT
END_METHOD

METHOD CALL_S010_READY
END_METHOD

METHOD CALL_S100_CLUTCH_CLOSE
END_METHOD

METHOD CALL_S200_SYNCHRON
END_METHOD

METHOD CALL_S300_CLUTCH_OPEN
END_METHOD

METHOD CALL_S998_ERROR
END_METHOD

(* ---- L_MB1P_COMCHANNELBASE.fb ---- *)
FUNCTION_BLOCK L_MB1P_COMCHANNELBASE EXTENDS L_MB1P_ComChannelSlaveBase
VAR_OUTPUT
	XMASTER : BOOL;
END_VAR
VAR_IN_OUT
	SCPAR : _scPar_TM_Base;
END_VAR
VAR
	ITFREFERENCECHECK2 : ITF_List;
	LISTFB : L_MB1P_ListControl := STRUCT(itfPar := THIS^);
	PPAR : POINTER TO _scPar_TM_MotionControl;
END_VAR
END_FUNCTION_BLOCK

METHOD CALL_ALLOCPOINTADR
END_METHOD

METHOD CALL_ERRORHANDLER
END_METHOD

METHOD CALL_RESETCOMMANDS
END_METHOD

METHOD CALL_RESETOUTPUTS
END_METHOD

(* ---- L_MB1P_COMCHANNELSLAVEBASE.fb ---- *)
FUNCTION_BLOCK L_MB1P_COMCHANNELSLAVEBASE
VAR_INPUT
	DATABUSIN : ITF_DataBus;
	XENABLE : BOOL;
	XPOINTERVALID : BOOL;
END_VAR
VAR_OUTPUT
	DATABUSOUT : ITF_DataBus := ComFB;
	XERROR : BOOL;
	EERRORID : L_IE1P_Error;
	XVALID : BOOL;
	XSLAVE : BOOL;
END_VAR
VAR
	COMFB : L_MB1P_Communication;
	PCOM : POINTER TO L_MB1P_Communication;
	PLIST_INT : POINTER TO L_MB1P_ListControl;
	ITFLIST : ITF_List;
	DATABUSIN_LOCK : ITF_DataBus;
	ITFREFERENCECHECK : ITF_DataBus;
	XENABLE_OLD : BOOL;
	PLIST : POINTER TO L_MB1P_ListControl;
	PPAR : POINTER TO _scPar_TM_MotionControl;
END_VAR
END_FUNCTION_BLOCK

METHOD CALL_ALLOCPOINTADR
END_METHOD

METHOD CALL_ERRORHANDLER
END_METHOD

METHOD CALL_OUTPUTS
END_METHOD

METHOD CALL_RESETCOMMANDS
END_METHOD

METHOD CALL_RESETOUTPUTS
END_METHOD

METHOD CALL_STATEMACHINE
END_METHOD

(* ---- L_MB1P_COMCHANNELSLAVESTATE.fb ---- *)
FUNCTION_BLOCK L_MB1P_COMCHANNELSLAVESTATE EXTENDS L_MB1P_ComChannelSlaveBase
VAR_OUTPUT
	XBUSY : BOOL;
	INUMOFELEMENTS : INT;
	IELEMENTNO : INT;
	IELEMENTID : INT;
	WCONNENCTIONTYPE : WORD;
END_VAR
VAR
	IELEMENTNO_LOCK : INT;
	ICALLNUM_LOCK : INT;
	PELEMENT_INT : POINTER TO L_MB1P_ChannelElement;
	XELEMENTVALID : BOOL;
	IIDNO : INT := 1;
	XCOMTOMASTERFAILED : BOOL;
	IDX : INT;
	PELEMENTLEFT : POINTER TO L_MB1P_ChannelElement;
	PELEMENTMASTER : POINTER TO L_MB1P_ChannelElement;
	PELEMENT : POINTER TO L_MB1P_ChannelElement;
END_VAR
END_FUNCTION_BLOCK

METHOD CALL_ALLOCPOINTADR
END_METHOD

METHOD CALL_ERRORHANDLER
END_METHOD

METHOD CALL_OUTPUTS
END_METHOD

METHOD CALL_RESETCOMMANDS
END_METHOD

METHOD CALL_RESETOUTPUTS
END_METHOD

METHOD CALL_STATEMACHINE
END_METHOD

(* ---- L_MB1P_COMCHANNELSTATE.fb ---- *)
FUNCTION_BLOCK L_MB1P_COMCHANNELSTATE EXTENDS L_MB1P_ComChannelBase
VAR_OUTPUT
	XBUSY : BOOL;
	INUMOFELEMENTS : INT;
	IELEMENTNO : INT;
	IELEMENTID : INT;
	WCONNENCTIONTYPE : WORD;
END_VAR
VAR
	IELEMENTNO_LOCK : INT;
	ICALLNUM_LOCK : INT;
	PELEMENT_INT : POINTER TO L_MB1P_ChannelElement;
	XELEMENTVALID : BOOL;
	IIDNO : INT := 1;
	XCOMTOMASTERFAILED : BOOL;
	IDX : INT;
	PELEMENTLEFT : POINTER TO L_MB1P_ChannelElement;
	PELEMENTMASTER : POINTER TO L_MB1P_ChannelElement;
	PELEMENT : POINTER TO L_MB1P_ChannelElement;
END_VAR
END_FUNCTION_BLOCK

METHOD CALL_ALLOCPOINTADR
END_METHOD

METHOD CALL_ERRORHANDLER
END_METHOD

METHOD CALL_OUTPUTS
END_METHOD

METHOD CALL_RESETCOMMANDS
END_METHOD

METHOD CALL_RESETOUTPUTS
END_METHOD

METHOD CALL_STATEMACHINE
END_METHOD

(* ---- L_MB1P_COMMUNICATION.fb ---- *)
FUNCTION_BLOCK L_MB1P_COMMUNICATION
VAR_INPUT
	ITFLIST : ITF_List;
	XLISTVALID : BOOL;
END_VAR
VAR
	PCOM : POINTER TO L_MB1P_Communication;
END_VAR
END_FUNCTION_BLOCK

(* ---- L_MB1P_DISTCORRECTIONWINDOW.fb ---- *)
FUNCTION_BLOCK L_MB1P_DISTCORRECTIONWINDOW
VAR_INPUT
	XENABLE : BOOL;
	XENABLEPOSITION : BOOL;
	LRCYCSETPOS : LREAL;
	LRCYCSETVEL : LREAL;
	XLOADSTARTPOS : BOOL;
	LRSTARTPOS : LREAL;
	XTPRECEIVEDIN : BOOL;
	LRSETCORRECTION : LREAL;
	XCORRWINDOWINXUNITS : BOOL;
	LRSETUPPERWINDOW : LREAL;
	LRSETLOWERWINDOW : LREAL;
	LRCYCPOSFEEDBACK : LREAL;
	DNSETNUMERATORAXISY : DWORD := 1;
	DNSETDENOMINATORAXISY : DWORD := 1;
	LRSETCYCLELENGTHX : LREAL;
	LRSETCYCLELENGTHY : LREAL;
END_VAR
VAR_OUTPUT
	XBUSY : BOOL;
	XCORRECTIONBUSY : BOOL;
	LRSETPOSOUT : LREAL;
	LRSETINTEGRATEDPOSITION : LREAL;
	LRSETPOSCORROUT : LREAL;
	LRSETPOSCORRRESIDUALOUT : LREAL;
	LRDELTAPOSCORROUT : LREAL;
	XCORRNEXTCYCLE : BOOL;
	XERROR : BOOL;
	EERRORID : L_IE1P_Error;
END_VAR
VAR
	LRDELTAPOSTOTAL : LREAL;
	LRMASTERDISTANCE : LREAL;
	LRPOSITIONSET : LREAL;
	LRPOSITIONNORMED : LREAL;
	LRPOSITIONOUTNORMED : LREAL;
	LRDELTAPOSCORRECTION : LREAL;
	LRPOSITIONSETOLD : LREAL;
	LRPOSITIONSETAXISOUT : LREAL;
	BYSTEPPER : BYTE;
	LRCORRECTIONDISTANCELOCAL : LREAL;
	LRCORRECTIONLOCAL : LREAL;
	L_DIFFERENTIATE : L_MC2P_Differentiate;
	INTEGRATOR : L_MC1P_IntegrateAxis;
	LRDELTAPOSOUT : LREAL;
	XEXECUTECORRECTIONINTERN : BOOL;
	XPOSITIVEDIRECTION : BOOL := FALSE;
	LRCORRECTIONDISTANCE : LREAL;
	LRUPPERWINDOWINTERNAL : LREAL;
	LRLOWERWINDOWINTERNAL : LREAL;
	LRTASKCYCLE : LREAL;
	XCORRECTIONACTIVE : BOOL;
	LRCORRECTIONLOCAL1 : LREAL;
	XTPRECEIVEDOLD : BOOL;
	LRINTEGRATORSPEED : LREAL;
	XWINDOWINCYCLE : BOOL;
	LRDELTAWINDOW : LREAL;
	LRCYCPOSINTOOLINTERNAL : LREAL;
	LRUPPERWINDOWINTERNALDELTA : LREAL;
	LRLOWERWINDOWINTERNALDELTA : LREAL;
	XINIT : BOOL := TRUE;
	XINITOUTOFCORRWINDOW : BOOL := TRUE;
	LRLOWERWINDOWINTERNALOLD : LREAL;
	LRUPPERWINDOWINTERNALOLD : LREAL;
	LRCYCPOSFEEDBACKINT : LREAL;
	XCORRECTIONBUSYOLD : BOOL;
	LRSETPOSCORROUTOLD : LREAL;
	LRCYCPOSINTOOLINTERNAL_CASE : LREAL;
	XWINDOWCHANGEDFLAG : BOOL := FALSE;
	LRCYCLELENGTH_INT : LREAL;
	LROFFSET_INT : LREAL;
	LRCYCPOSINTOOLINTERNAL_0LD : LREAL;
	LRPOSITIONNORMED_OLD : LREAL;
	LRPOSITIONNORMED_DIF : LREAL;
	XPOSCORR : BOOL;
	XTPSTORED_INT : BOOL;
	LRSETCORRECTIONSTORED_INT : LREAL;
	XINCORRWINDOW : BOOL;
	XINCORRWINDOWOLD : BOOL;
	LRSETPOSOUTCOMP : LREAL;
	LRCYCPOSINTOOLINTERNALOLD : LREAL;
	LRDELTAPOSOUTINTERNAL : LREAL;
	BYSTEPPEROLD : BYTE := 0;
END_VAR
END_FUNCTION_BLOCK

(* ---- L_MB1P_GEARBOXPOSITION.fb ---- *)
FUNCTION_BLOCK L_MB1P_GEARBOXPOSITION EXTENDS L_MB1P_GearboxPositionBase
VAR_IN_OUT
	AXISX : AXIS_REF;
	AXISY : AXIS_REF;
END_VAR
END_FUNCTION_BLOCK

METHOD CALL_ERRORHANDLER
END_METHOD

(* ---- L_MB1P_GEARBOXPOSITIONBASE.fb ---- *)
FUNCTION_BLOCK L_MB1P_GEARBOXPOSITIONBASE
VAR_INPUT
	XENABLE : BOOL;
	LRPOSX : LREAL;
	DWNUMERATOR : DWORD := 1;
	DWDENOMINATOR : DWORD := 1;
	XLOADPOSY : BOOL;
	LRLOADPOSY : LREAL;
	LNLOADPOSYRESIDUAL : LINT;
END_VAR
VAR_OUTPUT
	LRPOSY : LREAL;
	LNACTPOSYRESIDUAL : LINT;
	XERROR : BOOL := FALSE;
	EERRORID : L_IE1P_Error := 0;
END_VAR
VAR
	XINIT : BOOL := FALSE;
	LNPOSX : LINT := 0;
	LNPOSY : LINT := 0;
	LNPOSXOLD : LINT := 0;
	LNPOSXDIFF : LINT := 0;
	LNPOSYDIFF : LINT := 0;
	LNPOSYOLD : LINT := 0;
	LNRES_GEARBOX : LINT := 0;
	LRLENX : LREAL;
	LRLENY : LREAL;
	LRLENXOLD : LREAL;
	LRLENYOLD : LREAL;
END_VAR
END_FUNCTION_BLOCK

METHOD CALL_S000_CYCLIC
END_METHOD

METHOD CALL_ERRORHANDLER
END_METHOD

METHOD CALL_RESET
END_METHOD

METHOD L_HLPMODULOADD : LREAL
VAR_INPUT
	LRINPUT : LINT;
	LROFFSET : LINT;
	LRLENGHT : LINT;
END_VAR
END_METHOD

METHOD L_HLPMODULODIFF : LREAL
VAR_INPUT
	LRDIFF : LINT;
	LRLEN : LINT;
END_VAR
END_METHOD

METHOD L_HLPMULDIV : LREAL
VAR_INPUT
	LNINPUT : LINT;
	DWNUMERATOR : DWORD;
	DWDENOMINATOR : DWORD;
	PLNRES : POINTER TO LINT;
END_VAR
END_METHOD

(* ---- L_MB1P_GEARBOXPOSITIONINPUT.fb ---- *)
FUNCTION_BLOCK L_MB1P_GEARBOXPOSITIONINPUT EXTENDS L_MB1P_GearboxPositionBase
VAR_INPUT
	LRCYCLELENGTHX : LREAL;
	LRCYCLELENGTHY : LREAL;
END_VAR
END_FUNCTION_BLOCK

(* ---- L_MB1P_GENERATETPTIMESTAMP.fb ---- *)
FUNCTION_BLOCK L_MB1P_GENERATETPTIMESTAMP
VAR_INPUT
	XENABLE : BOOL;
	XTPRECEIVED : BOOL;
	LRACTTPPOSIN : LREAL;
	LRCYCPOSTPAXIS : LREAL;
	LRCYCLELENGTHTPAXIS : LREAL;
	LRCYCLELENGTHTARGETAXIS : LREAL;
	LRTASKCYCLELENGTH : LREAL;
END_VAR
VAR_OUTPUT
	XTPRECEIVEDOUT : BOOL;
	LRTPACTTIMESTAMP : LREAL;
	XERROR : BOOL;
END_VAR
VAR
	LRPOSFIFOX : ARRAY [1..20] OF LREAL := [10(0)];
	LRPOSFIFOREG : ARRAY [1..20] OF LREAL := [10(0)];
	BYCOUNTER : INT := 1;
	LRSTACKDIFFERENCE : LREAL;
	LRTPDELTAINMS : LREAL;
	LRDELTAPCT : LREAL;
	XTPRECEIVEDOLD : BOOL;
	LRTEMP : LREAL;
	IDIRECTION : INT;
	LRACTTPPOSINOLD : LREAL;
END_VAR
END_FUNCTION_BLOCK

METHOD SEARCHINSTACKNEGATIVE
END_METHOD

METHOD SEARCHINSTACKPOSITIVE
END_METHOD

(* ---- L_MB1P_HLPRAMPGENERATOR.fb ---- *)
FUNCTION_BLOCK L_MB1P_HLPRAMPGENERATOR
VAR_INPUT
	LRACC : LREAL;
	LRDEC : LREAL;
	LRVEL : LREAL;
	LRJERKACC : LREAL;
	LRJERKDEC : LREAL;
	LRTASKCYCLE : LREAL;
END_VAR
VAR_OUTPUT
	LRSETVEL : LREAL;
	LRSETACCDEC : LREAL;
	DNSTATE : DINT;
END_VAR
VAR
	ALRACCLIMIT : ARRAY [0..1] OF LREAL;
	ALRJERKABS : ARRAY [0..1] OF LREAL;
	LRVELINTERNAL : LREAL;
	DWINDEX : DWORD;
	LRVELDIFF : LREAL;
	LRVELCOMPARE : LREAL;
	LRACCINTERNAL : LREAL;
	C_RG_ACC : WORD := 0;
	C_RG_DEC : WORD := 1;
	C_RG_MINJERK : LREAL := 1;
	C_RG_STATE_INI : DINT := 0;
	C_RG_STATE_CNS : DINT := 1;
	C_RG_STATE_ACC : DINT := 2;
	C_RG_STATE_DEC : DINT := 3;
END_VAR
END_FUNCTION_BLOCK

METHOD RG_GETDEC : BOOL
VAR_INPUT
	LRVELDIFF : LREAL;
	LRVEL : LREAL;
END_VAR
END_METHOD

METHOD RG_MAXJERKINDEX : WORD
VAR_INPUT
	VAR1 : LREAL;
	VAR2 : LREAL;
	IND1 : WORD;
	IND2 : WORD;
END_VAR
END_METHOD

METHOD RG_REDACC : BOOL
VAR_INPUT
	LRVELDIFF : LREAL;
	LRACC : LREAL;
END_VAR
END_METHOD

METHOD SETSTARTVALUES
VAR_INPUT
	LRVEL : LREAL;
	LRACC : LREAL;
END_VAR
END_METHOD

METHOD TFM_RG_CALCDELTAVEL
END_METHOD

METHOD TFM_RG_CALCJERK : LREAL
VAR_INPUT
	VEL : LREAL;
	ACC : LREAL;
END_VAR
END_METHOD

METHOD TFM_RG_CALCPARAMETER
END_METHOD

METHOD TFM_RG_REDACC
END_METHOD

METHOD TFM_RG_VELDIFFNEG
END_METHOD

METHOD TFM_RG_VELDIFFPOS
END_METHOD

METHOD TFM_RG_VELTARGET
END_METHOD

(* ---- L_MB1P_LISTCONTROL.fb ---- *)
FUNCTION_BLOCK L_MB1P_LISTCONTROL
VAR_OUTPUT
	XERROR : BOOL;
	EERRORID : L_IE1P_Error;
	XLOCK : BOOL;
	XLISTVALID : BOOL;
	IFILLSTATE : INT;
	IELEMENTFIRST : INT;
	IELEMENTLAST : INT;
	ITFPAR : ITF_DataBusPar;
END_VAR
VAR
	DWID : __XWORD;
	XINITDONE : BOOL := FALSE;
	ARSCELEMENT : ARRAY [1..c_iElementNum] OF L_MB1P_ChannelElement;
	ASCDATA : ARRAY [1..c_iElementNum] OF L_MB1P_ChannelData;
	SCHEADDATA : L_MB1P_ChannelHeadData;
	ISTOREINSERELEMENTID : INT;
	IDX : INT;
	C_IELEMENTNUM : INT := 10;
	PLIST : POINTER TO L_MB1P_ListControl;
	PPAR : POINTER TO _scPar_TM_MotionControl;
END_VAR
END_FUNCTION_BLOCK

METHOD DELETELISTELEMENTID : BOOL
VAR_IN_OUT
	IIDNO : INT;
END_VAR
END_METHOD

METHOD DISABLE : BOOL
END_METHOD

METHOD GETELEMENTFIRST : POINTER TO L_MB1P_ChannelElement
VAR_OUTPUT
	XELEMENTVALID : BOOL;
	PELEMENT : POINTER TO L_MB1P_ChannelElement;
	IIDNO : INT;
	IELEMENTNO : INT;
END_VAR
END_METHOD

METHOD GETELEMENTID : POINTER TO L_MB1P_ChannelElement
VAR_OUTPUT
	XELEMENTVALID : BOOL;
	PELEMENT : POINTER TO L_MB1P_ChannelElement;
	IELEMENTNO : INT;
END_VAR
VAR_IN_OUT
	IIDNO : INT;
END_VAR
END_METHOD

METHOD GETELEMENTLAST : POINTER TO L_MB1P_ChannelElement
VAR_OUTPUT
	XELEMENTVALID : BOOL;
	PELEMENT : POINTER TO L_MB1P_ChannelElement;
	IIDNO : INT;
	IELEMENTNO : INT;
END_VAR
END_METHOD

METHOD GETELEMENTNO : POINTER TO L_MB1P_ChannelElement
VAR_OUTPUT
	XELEMENTVALID : BOOL;
	PELEMENT : POINTER TO L_MB1P_ChannelElement;
	IIDNO : INT;
END_VAR
VAR_IN_OUT
	IELEMENTNO : INT;
END_VAR
END_METHOD

METHOD GETENDELEMENT : POINTER TO L_MB1P_ChannelElement
VAR_OUTPUT
	XELEMENTVALID : BOOL;
	PELEMENT : POINTER TO L_MB1P_ChannelElement;
	IIDNO : INT;
	IELEMENTNO : INT;
END_VAR
END_METHOD

METHOD GETID : __XWORD
END_METHOD

METHOD GETSTARTELEMENT : POINTER TO L_MB1P_ChannelElement
VAR_OUTPUT
	XELEMENTVALID : BOOL;
	PELEMENT : POINTER TO L_MB1P_ChannelElement;
	IIDNO : INT;
	IELEMENTNO : INT;
END_VAR
END_METHOD

METHOD GETPDATA : __XWORD
VAR_INPUT
	IIDNO : INT;
END_VAR
END_METHOD

METHOD GETPELEMENTLEFT : POINTER TO L_MB1P_ChannelElement
VAR_IN_OUT
	IIDNO : INT;
END_VAR
END_METHOD

METHOD GETPELEMENTRIGHT : POINTER TO L_MB1P_ChannelElement
VAR_IN_OUT
	IIDNO : INT;
END_VAR
END_METHOD

METHOD GETPHEADDATA : __XWORD
END_METHOD

METHOD INIT : BOOL
END_METHOD

METHOD INITDATA
VAR_IN_OUT
	IIDNO : INT;
END_VAR
END_METHOD

METHOD INSERTELEMENTAFTERELEMENTID : POINTER TO L_MB1P_ChannelElement
VAR_INPUT
	IIDNOLEFT : INT;
END_VAR
VAR_OUTPUT
	XELEMENTVALID : BOOL;
	PELEMENT : POINTER TO L_MB1P_ChannelElement;
	IIDNO : INT := 1;
	IELEMENTNO : INT;
END_VAR
END_METHOD

METHOD INSERTELEMENTAFTERELEMENTNO : POINTER TO L_MB1P_ChannelElement
VAR_INPUT
	IELEMENTNOLEFT : INT;
END_VAR
VAR_OUTPUT
	XELEMENTVALID : BOOL;
	PELEMENT : POINTER TO L_MB1P_ChannelElement;
	IIDNO : INT := 1;
	IELEMENTNO : INT;
END_VAR
END_METHOD

METHOD INSERTNEWELEMENT : POINTER TO L_MB1P_ChannelElement
VAR_OUTPUT
	XELEMENTVALID : BOOL;
	PELEMENT : POINTER TO L_MB1P_ChannelElement;
	IIDNO : INT := 1;
	IELEMENTNO : INT;
END_VAR
END_METHOD

METHOD LOCK : BOOL
END_METHOD

METHOD SETERROR : BOOL
VAR_INPUT
	EERRID : L_IE1P_Error;
END_VAR
END_METHOD

METHOD UNLOCK : BOOL
END_METHOD

(* ---- L_MB1P_MARKREGISTER.fb ---- *)
FUNCTION_BLOCK L_MB1P_MARKREGISTER
VAR_INPUT
	XENABLE : BOOL;
	LRCYCSETVEL : LREAL;
	XTPRECEIVEDIN : BOOL;
	LRSETTPDIFFERENCE : LREAL;
	LRMARKSTACKLENGTH : LREAL;
	XCORRECTIONBUSY : BOOL;
	LRSETPOSCORRIN : LREAL;
END_VAR
VAR_OUTPUT
	XTPRECEIVEDOUT : BOOL;
	LRTPDIFFERENCEOUT : LREAL;
	LRTOTALSTACKDIFFERENCEOUT : LREAL;
	XERROR : BOOL := FALSE;
	EERRORID : L_IE1P_Error;
END_VAR
VAR
	LRTPDIFFERENCES : ARRAY [1..64] OF LREAL := [64(0)];
	LRTPPOSITION : ARRAY [1..64] OF LREAL := [64(0)];
	XTPVALID : ARRAY [1..64] OF BOOL := [64(FALSE)];
	L_D94A_SDINTEGRATEAXIS1 : L_MC1P_IntegrateAxis;
	COUNTERIN : WORD := 1;
	COUNTEROUT : WORD := 1;
	DWINTEGRATORVALUE : DWORD := 0;
	LRINTEGRATORPOS : LREAL := 0;
	LRTASKCYCLE : LREAL;
	LRPOSDIFF : LREAL;
	LRPOSTOREGISTEREND : LREAL;
	XREGISTERFULL : BOOL;
	LRPOSDIFFINSTACK : LREAL := 0;
	DWCOUNTER : DWORD;
	XINIT : BOOL;
	XWAITINGFORCORRECTIONDONE : BOOL;
	XCORRETIONSTARTED : BOOL;
	LRACTUALTPDIFFERENCE : LREAL;
	XCORRECTIONBUSY_OLD : BOOL;
	LRSETPOSCORRIN_OLD : LREAL;
END_VAR
END_FUNCTION_BLOCK

METHOD CALL_CALCULATETOTALSTACK
END_METHOD

METHOD CALL_WAITFORCORRECTION
END_METHOD

(* ---- L_MB1P_MARKSTACK.fb ---- *)
FUNCTION_BLOCK L_MB1P_MARKSTACK
VAR_INPUT
	XENABLE : BOOL;
	XTPRECEIVEDIN : BOOL;
	LRACTTPPOSITION : LREAL;
	LRACTVELMATERIAL : LREAL;
	LRACTPOSITIONTPAXIS : LREAL;
	LRCYCLELENGTHTPAXIS : LREAL;
	LRMARKSTACKLENGTH : LREAL;
END_VAR
VAR_OUTPUT
	XTPRECEIVEDOUT : BOOL;
	LRACTTPPOSITIONOUT : LREAL;
	XERROR : BOOL := FALSE;
	EERRORID : WORD;
	LRTPDIFFOUT : LREAL;
END_VAR
VAR
	ALRINTEGRATORSTARTPOS : ARRAY [1..64] OF LREAL := [64(0)];
	ALRINTEGRATORDIST : ARRAY [1..64] OF LREAL := [64(0)];
	ALRLASTSCAN : ARRAY [1..64] OF LREAL := [64(0)];
	XTPVALID : ARRAY [1..64] OF BOOL := [64(FALSE)];
	XREGISTERFULL : BOOL := FALSE;
	XINIT : BOOL := TRUE;
	WCOUNTER : WORD;
	WCOUNTERIN : WORD := 1;
	WCOUNTEROUT : WORD := 1;
	LRINTEGRATORPOS : LREAL := 0;
	LRTASKCYCLE : LREAL;
	LRCYCPOSDIFF : LREAL := 0;
	LRPOSTOREGISTEREND : LREAL := 0;
	XTPRECEIVEDINOLD : BOOL;
	LRMARKSTACKLENGTHOLD : LREAL;
	LRACTPOSITIONTPAXISCOMP : LREAL;
END_VAR
END_FUNCTION_BLOCK

METHOD CALL_INITMARKSTACK
END_METHOD

(* ---- L_MB1P_MARKWINDOW.fb ---- *)
FUNCTION_BLOCK L_MB1P_MARKWINDOW
VAR_INPUT
	XENABLE : BOOL;
	LRCYCREGISTERPOS : LREAL;
	LRCYCSETVEL : LREAL;
	XTPRECEIVEDIN : BOOL;
	LRACTTPPOSIN : LREAL;
	XTEACHMARKWINDOW : BOOL;
	LRSETMARKDISTANCE : LREAL;
	LRMARKSENSORPOSITION : LREAL;
	LRSETMARKWINDOW : LREAL;
	LRSETOFFSETMARKWINDOW : LREAL;
	DWMAXTPNOTDETECTED : DWORD;
END_VAR
VAR_OUTPUT
	XTPRECEIVEDOUT : BOOL;
	XTPWINDOWOPEN : BOOL;
	XTPWINDOWOPENCOMP : BOOL;
	LRTPDELTAPOSCOMP : LREAL;
	XTPINWINDOW : BOOL;
	XTPNOTINWINDOW : BOOL;
	XTPNOTDETECTED : BOOL;
	XTPSENSORTEACHED : BOOL;
	LRACTTPPOS : LREAL;
	XMAXTPNOTDETECTED : BOOL;
END_VAR
VAR
	XFIRSTSENSOR : BOOL;
	XTPWINDOWOPENOLD : BOOL;
	XTPNOTDETECTEDINTERNAL : BOOL;
	LRLOWERWINDOW : LREAL;
	LRUPPERWINDOW : LREAL;
	LRTPPOSINWINDOWTEST : LREAL;
	XTEACHTPSENSOROLD : BOOL;
	DWMISSEDTPCOUNTER : DWORD;
	LRACTUALREGISTERPOS : LREAL;
	XTPISINWINDOW : BOOL;
	XMISSEDTPDECREMENT : BOOL;
	LRDEADTIMEPOSDIFF : LREAL;
	LRUPPERWINDOWCOMP : LREAL;
	XTPCOMPWINDOWOPEN : BOOL;
	XTPCOMPWINDOWOPENOLD : BOOL := FALSE;
	LRLOWERWINDOWCOMP : LREAL;
	XTPRECEIVEDOLD : BOOL;
	LRACTUALREGISTERPOSOLD : LREAL;
	XTPRECEIVEDINTERNAL : BOOL;
	LRTASKCYCLE : LREAL;
END_VAR
END_FUNCTION_BLOCK

(* ---- L_MB1P_MARKWINDOWRELATIVE.fb ---- *)
FUNCTION_BLOCK L_MB1P_MARKWINDOWRELATIVE
VAR_INPUT
	XENABLE : BOOL;
	LRTPWINDOWSIZE : LREAL;
	LRCYCVEL : LREAL;
	XTPRECEIVE : BOOL;
	LRACTTPPOSIN : LREAL;
	LRCYCLELENGTH : LREAL;
	XTEACHMARKWINDOW : BOOL;
	LRSETOFFSETTPWINDOW : LREAL;
	DWMAXTPNOTDETECTED : DWORD;
	LRSTARTPOSITION : LREAL;
END_VAR
VAR_OUTPUT
	XTPRECEIVED : BOOL;
	XTPWINDOWOPEN : BOOL;
	XTPWINDOWOPENCOMP : BOOL;
	LRTPDELTAPOSCOMP : LREAL;
	XTPINWINDOW : BOOL;
	XTPNOTINWINDOW : BOOL;
	XTPNOTDETECTED : BOOL;
	XTPSENSORTEACHED : BOOL;
	LRACTTPPOS : LREAL;
	XMAXTPNOTDETECTED : BOOL;
END_VAR
VAR
	LRMARKWINDOWINTEGRATOROLD : LREAL;
	XFIRSTSENSOR : BOOL;
	XTPWINDOWOPENOLD : BOOL;
	XTPNOTDETECTEDINTERNAL : BOOL;
	LRLOWERWINDOW : LREAL;
	LRUPPERWINDOW : LREAL;
	LRTPPOSINWINDOWTEST : LREAL;
	XTEACHTPSENSOROLD : BOOL;
	DWMISSEDTPCOUNTER : DWORD;
	LRACTUALREGISTERPOS : LREAL;
	XTPISINWINDOW : BOOL;
	XMISSEDTPDECREMENT : BOOL;
	LRDEADTIMEPOSDIFF : LREAL;
	LRUPPERWINDOWCOMP : LREAL;
	XTPCOMPWINDOWOPEN : BOOL;
	XTPCOMPWINDOWOPENOLD : BOOL := FALSE;
	LRLOWERWINDOWCOMP : LREAL;
	XTPRECEIVEDOLD : BOOL;
	LRACTUALREGISTERPOSOLD : LREAL;
	XTPRECEIVEDINTERNAL : BOOL;
	LRTASKCYCLE : LREAL;
	LRTPWINDOWSIZE_INT : LREAL;
	LRMARKWINDOWINTEGRATOR : LREAL := 0;
	LRDEADTIMETP : LREAL;
	LRACTUALTPPOSITION : LREAL;
END_VAR
END_FUNCTION_BLOCK

(* ---- L_MB1P_MATERIALCOUNTER.fb ---- *)
FUNCTION_BLOCK L_MB1P_MATERIALCOUNTER
VAR_INPUT
	XENABLE : BOOL;
	LRPOSIN : LREAL;
	LRACTVELIN : LREAL;
	LRTASKCYCLE : LREAL;
	LRPOSINSLAVE : LREAL;
	LRCYCLELEN : LREAL;
	XLOADSTARTPOS : BOOL;
	XSETMATERIALCOUNTER : BOOL;
	LRSETMATERIALPOS : LREAL;
	XLOADDELTAPOS : BOOL;
	LRSETDELTAPOS : LREAL;
	XSTARTFLYINGSAW : BOOL;
END_VAR
VAR_OUTPUT
	LNMATERIALPOS_E8 : LINT;
	LNMATERIALPOSOUT_E8 : LINT;
	LRMATERIALCOUNTER : LREAL;
	LRDELTAMATERIALPOS : LREAL;
END_VAR
VAR_IN_OUT
	AXIS : AXIS_REF;
END_VAR
VAR
	LNMODULOPOS_E8 : LINT;
	LNMODULOPOSOLD_E8 : LINT;
	LNCYCLELEN_E8 : LINT;
	LNPOSXDIFF : LINT;
	LNLENX_INT : LINT;
	LNMATERIALPOS_E8_OLD : LINT;
	LNDELTAMATERIALPOS : LINT;
	XSETMATERIALCOUNTER_OLD : BOOL;
	XINITDONE : BOOL;
	LROFFSET : LREAL;
	PAXIS : POINTER TO _AXIS_REF_REAL;
	LRJITTERPOS : LREAL;
	LNJITTERPOS : LINT;
	XENABLE_OLD : BOOL;
END_VAR
END_FUNCTION_BLOCK

(* ---- L_MB1P_MATERIALLENGTHCOUNTERFROMPOS.fb ---- *)
FUNCTION_BLOCK L_MB1P_MATERIALLENGTHCOUNTERFROMPOS
VAR_INPUT
	XENABLE : BOOL;
	LRACTPOSIN : LREAL;
	WFILTERDEPTH : WORD := 0;
	LRCYCLELENGTH : LREAL := 360;
	LRSETFEEDCONSTANT : LREAL := 360;
	XSETMATERIALCOUNTER : BOOL;
	LRSETMATERIALPOS : LREAL;
END_VAR
VAR_OUTPUT
	XBUSY : BOOL;
	XERROR : BOOL;
	EERRORID : L_IE1P_Error;
	LRMATERIALCOUNTER : LREAL;
	LRREVCOUNTER : LREAL;
	LIREVCOUNTER : LINT;
	LIREVCOUNTERMID : LINT;
	LRREVCOUNTERRESIDUAL : LREAL;
END_VAR
VAR_IN_OUT
	LIREVCOUNTERRETAIN : LINT;
	LRREVCOUNTERRESIDUALRETAIN : LREAL;
END_VAR
VAR
	WSTATE : WORD;
	XENABLE_OLD : BOOL;
	XSETMATERIALCOUNTER_OLD : BOOL;
	LRSTARTPOS_INT : LREAL;
	LRACTPOSIN_INT : LREAL;
	LIREVCOUNTER_OLD : LINT;
	LRREVCOUNTER_INT : LREAL;
	LIREVCOUNTERMID_OLD : LINT;
	LRREVCOUNTERMID_INT : LREAL;
	XERRORRECIVEDLIMIT : BOOL;
	LRREVCOUNTERRESIDUAL_OFFSET : LREAL;
	LRACTPOSIN_OLD : LREAL;
	C_LRLINTMAXVALUEPOS : LREAL := 2#111111111111111111111111111111111111111111111111111111111111111;
	C_LRLINTMAXVALUENEG : LREAL := -2#111111111111111111111111111111111111111111111111111111111111111;
END_VAR
END_FUNCTION_BLOCK

METHOD CALL_CALCMATERAILCOUNTER
END_METHOD

METHOD CALL_ERRORHANDLER
END_METHOD

METHOD CALL_OUTPUT
END_METHOD

METHOD CALL_RESETCOMMANDS
END_METHOD

METHOD CALL_RESETOUTPUT
END_METHOD

(* ---- L_MB1P_MATERIALLENGTHCOUNTERFROMVEL.fb ---- *)
FUNCTION_BLOCK L_MB1P_MATERIALLENGTHCOUNTERFROMVEL
VAR_INPUT
	XENABLE : BOOL;
	LRACTVELIN : LREAL;
	RFILTERTIME : REAL := 0.0;
	XSETMATERIALCOUNTER : BOOL;
	LRSETMATERIALPOS : LREAL;
END_VAR
VAR_OUTPUT
	XBUSY : BOOL;
	XWARNING : BOOL;
	EERRORID : L_IE1P_Error;
	LRMATERIALCOUNTER : LREAL;
END_VAR
VAR_IN_OUT
	LRSETMATERIALPOSRETAIN : LREAL;
END_VAR
VAR
	WSTATE : WORD;
	XENABLE_OLD : BOOL;
	XSETMATERIALCOUNTER_OLD : BOOL;
	LRTASKCYCLE : LREAL;
	LIPOS_INT : LINT;
	LIDELTAPOS_INT : LINT;
	LIPOS_OLD : LINT;
	LIIDX : LINT;
	LRMATERIALCOUNTERCOUNTER_INT : LREAL;
	LRMATERIALOFFSET_INT : LREAL;
	FB_PT1FILTER : L_USPP_PT1Filter;
END_VAR
END_FUNCTION_BLOCK

METHOD CALL_CALCMATERAILCOUNTER
END_METHOD

METHOD CALL_ERRORHANDLER
END_METHOD

METHOD CALL_FBMETHODS
END_METHOD

METHOD CALL_FB_PT1FILTER
END_METHOD

METHOD CALL_OUTPUT
END_METHOD

METHOD CALL_RESETCOMMANDS
END_METHOD

METHOD CALL_RESETOUTPUT
END_METHOD

METHOD CALL_STATEMACHINE
END_METHOD
